(* Logix 5000 project; controller TFF vendor 1 type 14 code 107 rev 34.11; software revision 34.03; part 11 of 36 *)

        [5,29].Action := -999, [5,29].Label := -999, [5,29].Criteria1Value := -1000000.0, [5,29].Criteria2Value := -1000000.0, [5,29].ActionValue := -1000000.0, [5,30].Criteria1 := -999, [5,30].Criteria1Operator := -999, [5,30].Boolean := -999, [5,30].Criteria2 := -999, [5,30].Criteria2Operator := -999, [5,30].Action := -999, [5,30].Label := -999, [5,30].Criteria1Value := -1000000.0, [5,30].Criteria2Value := -1000000.0, [5,30].ActionValue := -1000000.0, [5,31].Criteria1 := -999, [5,31].Criteria1Operator := -999, [5,31].Boolean := -999, [5,31].Criteria2 := -999, [5,31].Criteria2Operator := -999, [5,31].Action := -999, [5,31].Label := -999, [5,31].Criteria1Value := -1000000.0, [5,31].Criteria2Value := -1000000.0, [5,31].ActionValue := -1000000.0, [5,32].Criteria1 := -999, [5,32].Criteria1Operator := -999, [5,32].Boolean := -999, [5,32].Criteria2 := -999, [5,32].Criteria2Operator := -999, [5,32].Action := -999, [5,32].Label := -999, [5,32].Criteria1Value := -1000000.0, [5,32].Criteria2Value := -1000000.0, [5,32].ActionValue := -1000000.0, [5,33].Criteria1 := -999, [5,33].Criteria1Operator := -999, [5,33].Boolean := -999, [5,33].Criteria2 := -999, [5,33].Criteria2Operator := -999, [5,33].Action := -999, [5,33].Label := -999, [5,33].Criteria1Value := -1000000.0, [5,33].Criteria2Value := -1000000.0, [5,33].ActionValue := -1000000.0, [5,34].Criteria1 := -999, [5,34].Criteria1Operator := -999, [5,34].Boolean := -999, [5,34].Criteria2 := -999, [5,34].Criteria2Operator := -999, [5,34].Action := -999, [5,34].Label := -999, [5,34].Criteria1Value := -1000000.0, [5,34].Criteria2Value := -1000000.0, [5,34].ActionValue := -1000000.0, [5,35].Criteria1 := -999, [5,35].Criteria1Operator := -999, [5,35].Boolean := -999, [5,35].Criteria2 := -999, [5,35].Criteria2Operator := -999,
        [5,35].Action := -999, [5,35].Label := -999, [5,35].Criteria1Value := -1000000.0, [5,35].Criteria2Value := -1000000.0, [5,35].ActionValue := -1000000.0, [5,36].Criteria1 := -999, [5,36].Criteria1Operator := -999, [5,36].Boolean := -999, [5,36].Criteria2 := -999, [5,36].Criteria2Operator := -999, [5,36].Action := -999, [5,36].Label := -999, [5,36].Criteria1Value := -1000000.0, [5,36].Criteria2Value := -1000000.0, [5,36].ActionValue := -1000000.0, [5,37].Criteria1 := -999, [5,37].Criteria1Operator := -999, [5,37].Boolean := -999, [5,37].Criteria2 := -999, [5,37].Criteria2Operator := -999, [5,37].Action := -999, [5,37].Label := -999, [5,37].Criteria1Value := -1000000.0, [5,37].Criteria2Value := -1000000.0, [5,37].ActionValue := -1000000.0, [5,38].Criteria1 := -999, [5,38].Criteria1Operator := -999, [5,38].Boolean := -999, [5,38].Criteria2 := -999, [5,38].Criteria2Operator := -999, [5,38].Action := -999, [5,38].Label := -999, [5,38].Criteria1Value := -1000000.0, [5,38].Criteria2Value := -1000000.0, [5,38].ActionValue := -1000000.0, [5,39].Criteria1 := -999, [5,39].Criteria1Operator := -999, [5,39].Boolean := -999, [5,39].Criteria2 := -999, [5,39].Criteria2Operator := -999, [5,39].Action := -999, [5,39].Label := -999, [5,39].Criteria1Value := -1000000.0, [5,39].Criteria2Value := -1000000.0, [5,39].ActionValue := -1000000.0, [5,40].Criteria1 := -999, [5,40].Criteria1Operator := -999, [5,40].Boolean := -999, [5,40].Criteria2 := -999, [5,40].Criteria2Operator := -999, [5,40].Action := -999, [5,40].Label := -999, [5,40].Criteria1Value := -1000000.0, [5,40].Criteria2Value := -1000000.0, [5,40].ActionValue := -1000000.0, [5,41].Criteria1 := -999, [5,41].Criteria1Operator := -999, [5,41].Boolean := -999, [5,41].Criteria2 := -999, [5,41].Criteria2Operator := -999,
        [5,41].Action := -999, [5,41].Label := -999, [5,41].Criteria1Value := -1000000.0, [5,41].Criteria2Value := -1000000.0, [5,41].ActionValue := -1000000.0, [5,42].Criteria1 := -999, [5,42].Criteria1Operator := -999, [5,42].Boolean := -999, [5,42].Criteria2 := -999, [5,42].Criteria2Operator := -999, [5,42].Action := -999, [5,42].Label := -999, [5,42].Criteria1Value := -1000000.0, [5,42].Criteria2Value := -1000000.0, [5,42].ActionValue := -1000000.0, [5,43].Criteria1 := -999, [5,43].Criteria1Operator := -999, [5,43].Boolean := -999, [5,43].Criteria2 := -999, [5,43].Criteria2Operator := -999, [5,43].Action := -999, [5,43].Label := -999, [5,43].Criteria1Value := -1000000.0, [5,43].Criteria2Value := -1000000.0, [5,43].ActionValue := -1000000.0, [5,44].Criteria1 := -999, [5,44].Criteria1Operator := -999, [5,44].Boolean := -999, [5,44].Criteria2 := -999, [5,44].Criteria2Operator := -999, [5,44].Action := -999, [5,44].Label := -999, [5,44].Criteria1Value := -1000000.0, [5,44].Criteria2Value := -1000000.0, [5,44].ActionValue := -1000000.0, [5,45].Criteria1 := -999, [5,45].Criteria1Operator := -999, [5,45].Boolean := -999, [5,45].Criteria2 := -999, [5,45].Criteria2Operator := -999, [5,45].Action := -999, [5,45].Label := -999, [5,45].Criteria1Value := -1000000.0, [5,45].Criteria2Value := -1000000.0, [5,45].ActionValue := -1000000.0, [5,46].Criteria1 := -999, [5,46].Criteria1Operator := -999, [5,46].Boolean := -999, [5,46].Criteria2 := -999, [5,46].Criteria2Operator := -999, [5,46].Action := -999, [5,46].Label := -999, [5,46].Criteria1Value := -1000000.0, [5,46].Criteria2Value := -1000000.0, [5,46].ActionValue := -1000000.0, [5,47].Criteria1 := -999, [5,47].Criteria1Operator := -999, [5,47].Boolean := -999, [5,47].Criteria2 := -999, [5,47].Criteria2Operator := -999,
        [5,47].Action := -999, [5,47].Label := -999, [5,47].Criteria1Value := -1000000.0, [5,47].Criteria2Value := -1000000.0, [5,47].ActionValue := -1000000.0, [5,48].Criteria1 := -999, [5,48].Criteria1Operator := -999, [5,48].Boolean := -999, [5,48].Criteria2 := -999, [5,48].Criteria2Operator := -999, [5,48].Action := -999, [5,48].Label := -999, [5,48].Criteria1Value := -1000000.0, [5,48].Criteria2Value := -1000000.0, [5,48].ActionValue := -1000000.0, [5,49].Criteria1 := -999, [5,49].Criteria1Operator := -999, [5,49].Boolean := -999, [5,49].Criteria2 := -999, [5,49].Criteria2Operator := -999, [5,49].Action := -999, [5,49].Label := -999, [5,49].Criteria1Value := -1000000.0, [5,49].Criteria2Value := -1000000.0, [5,49].ActionValue := -1000000.0, [5,50].Criteria1 := -999, [5,50].Criteria1Operator := -999, [5,50].Boolean := -999, [5,50].Criteria2 := -999, [5,50].Criteria2Operator := -999, [5,50].Action := -999, [5,50].Label := -999, [5,50].Criteria1Value := -1000000.0, [5,50].Criteria2Value := -1000000.0, [5,50].ActionValue := -1000000.0, [5,51].Criteria1 := -999, [5,51].Criteria1Operator := -999, [5,51].Boolean := -999, [5,51].Criteria2 := -999, [5,51].Criteria2Operator := -999, [5,51].Action := -999, [5,51].Label := -999, [5,51].Criteria1Value := -1000000.0, [5,51].Criteria2Value := -1000000.0, [5,51].ActionValue := -1000000.0, [5,52].Criteria1 := -999, [5,52].Criteria1Operator := -999, [5,52].Boolean := -999, [5,52].Criteria2 := -999, [5,52].Criteria2Operator := -999, [5,52].Action := -999, [5,52].Label := -999, [5,52].Criteria1Value := -1000000.0, [5,52].Criteria2Value := -1000000.0, [5,52].ActionValue := -1000000.0, [5,53].Criteria1 := -999, [5,53].Criteria1Operator := -999, [5,53].Boolean := -999, [5,53].Criteria2 := -999, [5,53].Criteria2Operator := -999,
        [5,53].Action := -999, [5,53].Label := -999, [5,53].Criteria1Value := -1000000.0, [5,53].Criteria2Value := -1000000.0, [5,53].ActionValue := -1000000.0, [5,54].Criteria1 := -999, [5,54].Criteria1Operator := -999, [5,54].Boolean := -999, [5,54].Criteria2 := -999, [5,54].Criteria2Operator := -999, [5,54].Action := -999, [5,54].Label := -999, [5,54].Criteria1Value := -1000000.0, [5,54].Criteria2Value := -1000000.0, [5,54].ActionValue := -1000000.0, [5,55].Criteria1 := -999, [5,55].Criteria1Operator := -999, [5,55].Boolean := -999, [5,55].Criteria2 := -999, [5,55].Criteria2Operator := -999, [5,55].Action := -999, [5,55].Label := -999, [5,55].Criteria1Value := -1000000.0, [5,55].Criteria2Value := -1000000.0, [5,55].ActionValue := -1000000.0, [5,56].Criteria1 := -999, [5,56].Criteria1Operator := -999, [5,56].Boolean := -999, [5,56].Criteria2 := -999, [5,56].Criteria2Operator := -999, [5,56].Action := -999, [5,56].Label := -999, [5,56].Criteria1Value := -1000000.0, [5,56].Criteria2Value := -1000000.0, [5,56].ActionValue := -1000000.0, [5,57].Criteria1 := -999, [5,57].Criteria1Operator := -999, [5,57].Boolean := -999, [5,57].Criteria2 := -999, [5,57].Criteria2Operator := -999, [5,57].Action := -999, [5,57].Label := -999, [5,57].Criteria1Value := -1000000.0, [5,57].Criteria2Value := -1000000.0, [5,57].ActionValue := -1000000.0, [5,58].Criteria1 := -999, [5,58].Criteria1Operator := -999, [5,58].Boolean := -999, [5,58].Criteria2 := -999, [5,58].Criteria2Operator := -999, [5,58].Action := -999, [5,58].Label := -999, [5,58].Criteria1Value := -1000000.0, [5,58].Criteria2Value := -1000000.0, [5,58].ActionValue := -1000000.0, [5,59].Criteria1 := -999, [5,59].Criteria1Operator := -999, [5,59].Boolean := -999, [5,59].Criteria2 := -999, [5,59].Criteria2Operator := -999,
        [5,59].Action := -999, [5,59].Label := -999, [5,59].Criteria1Value := -1000000.0, [5,59].Criteria2Value := -1000000.0, [5,59].ActionValue := -1000000.0, [5,60].Criteria1 := -999, [5,60].Criteria1Operator := -999, [5,60].Boolean := -999, [5,60].Criteria2 := -999, [5,60].Criteria2Operator := -999, [5,60].Action := -999, [5,60].Label := -999, [5,60].Criteria1Value := -1000000.0, [5,60].Criteria2Value := -1000000.0, [5,60].ActionValue := -1000000.0, [5,61].Criteria1 := -999, [5,61].Criteria1Operator := -999, [5,61].Boolean := -999, [5,61].Criteria2 := -999, [5,61].Criteria2Operator := -999, [5,61].Action := -999, [5,61].Label := -999, [5,61].Criteria1Value := -1000000.0, [5,61].Criteria2Value := -1000000.0, [5,61].ActionValue := -1000000.0, [5,62].Criteria1 := -999, [5,62].Criteria1Operator := -999, [5,62].Boolean := -999, [5,62].Criteria2 := -999, [5,62].Criteria2Operator := -999, [5,62].Action := -999, [5,62].Label := -999, [5,62].Criteria1Value := -1000000.0, [5,62].Criteria2Value := -1000000.0, [5,62].ActionValue := -1000000.0, [5,63].Criteria1 := -999, [5,63].Criteria1Operator := -999, [5,63].Boolean := -999, [5,63].Criteria2 := -999, [5,63].Criteria2Operator := -999, [5,63].Action := -999, [5,63].Label := -999, [5,63].Criteria1Value := -1000000.0, [5,63].Criteria2Value := -1000000.0, [5,63].ActionValue := -1000000.0, [5,64].Criteria1 := -999, [5,64].Criteria1Operator := -999, [5,64].Boolean := -999, [5,64].Criteria2 := -999, [5,64].Criteria2Operator := -999, [5,64].Action := -999, [5,64].Label := -999, [5,64].Criteria1Value := -1000000.0, [5,64].Criteria2Value := -1000000.0, [5,64].ActionValue := -1000000.0, [5,65].Criteria1 := -999, [5,65].Criteria1Operator := -999, [5,65].Boolean := -999, [5,65].Criteria2 := -999, [5,65].Criteria2Operator := -999,
        [5,65].Action := -999, [5,65].Label := -999, [5,65].Criteria1Value := -1000000.0, [5,65].Criteria2Value := -1000000.0, [5,65].ActionValue := -1000000.0, [5,66].Criteria1 := -999, [5,66].Criteria1Operator := -999, [5,66].Boolean := -999, [5,66].Criteria2 := -999, [5,66].Criteria2Operator := -999, [5,66].Action := -999, [5,66].Label := -999, [5,66].Criteria1Value := -1000000.0, [5,66].Criteria2Value := -1000000.0, [5,66].ActionValue := -1000000.0, [5,67].Criteria1 := -999, [5,67].Criteria1Operator := -999, [5,67].Boolean := -999, [5,67].Criteria2 := -999, [5,67].Criteria2Operator := -999, [5,67].Action := -999, [5,67].Label := -999, [5,67].Criteria1Value := -1000000.0, [5,67].Criteria2Value := -1000000.0, [5,67].ActionValue := -1000000.0, [5,68].Criteria1 := -999, [5,68].Criteria1Operator := -999, [5,68].Boolean := -999, [5,68].Criteria2 := -999, [5,68].Criteria2Operator := -999, [5,68].Action := -999, [5,68].Label := -999, [5,68].Criteria1Value := -1000000.0, [5,68].Criteria2Value := -1000000.0, [5,68].ActionValue := -1000000.0, [5,69].Criteria1 := -999, [5,69].Criteria1Operator := -999, [5,69].Boolean := -999, [5,69].Criteria2 := -999, [5,69].Criteria2Operator := -999, [5,69].Action := -999, [5,69].Label := -999, [5,69].Criteria1Value := -1000000.0, [5,69].Criteria2Value := -1000000.0, [5,69].ActionValue := -1000000.0, [5,70].Criteria1 := -999, [5,70].Criteria1Operator := -999, [5,70].Boolean := -999, [5,70].Criteria2 := -999, [5,70].Criteria2Operator := -999, [5,70].Action := -999, [5,70].Label := -999, [5,70].Criteria1Value := -1000000.0, [5,70].Criteria2Value := -1000000.0, [5,70].ActionValue := -1000000.0, [5,71].Criteria1 := -999, [5,71].Criteria1Operator := -999, [5,71].Boolean := -999, [5,71].Criteria2 := -999, [5,71].Criteria2Operator := -999,
        [5,71].Action := -999, [5,71].Label := -999, [5,71].Criteria1Value := -1000000.0, [5,71].Criteria2Value := -1000000.0, [5,71].ActionValue := -1000000.0, [5,72].Criteria1 := -999, [5,72].Criteria1Operator := -999, [5,72].Boolean := -999, [5,72].Criteria2 := -999, [5,72].Criteria2Operator := -999, [5,72].Action := -999, [5,72].Label := -999, [5,72].Criteria1Value := -1000000.0, [5,72].Criteria2Value := -1000000.0, [5,72].ActionValue := -1000000.0, [5,73].Criteria1 := -999, [5,73].Criteria1Operator := -999, [5,73].Boolean := -999, [5,73].Criteria2 := -999, [5,73].Criteria2Operator := -999, [5,73].Action := -999, [5,73].Label := -999, [5,73].Criteria1Value := -1000000.0, [5,73].Criteria2Value := -1000000.0, [5,73].ActionValue := -1000000.0, [5,74].Criteria1 := -999, [5,74].Criteria1Operator := -999, [5,74].Boolean := -999, [5,74].Criteria2 := -999, [5,74].Criteria2Operator := -999, [5,74].Action := -999, [5,74].Label := -999, [5,74].Criteria1Value := -1000000.0, [5,74].Criteria2Value := -1000000.0, [5,74].ActionValue := -1000000.0, [5,75].Criteria1 := -999, [5,75].Criteria1Operator := -999, [5,75].Boolean := -999, [5,75].Criteria2 := -999, [5,75].Criteria2Operator := -999, [5,75].Action := -999, [5,75].Label := -999, [5,75].Criteria1Value := -1000000.0, [5,75].Criteria2Value := -1000000.0, [5,75].ActionValue := -1000000.0, [5,76].Criteria1 := -999, [5,76].Criteria1Operator := -999, [5,76].Boolean := -999, [5,76].Criteria2 := -999, [5,76].Criteria2Operator := -999, [5,76].Action := -999, [5,76].Label := -999, [5,76].Criteria1Value := -1000000.0, [5,76].Criteria2Value := -1000000.0, [5,76].ActionValue := -1000000.0, [5,77].Criteria1 := -999, [5,77].Criteria1Operator := -999, [5,77].Boolean := -999, [5,77].Criteria2 := -999, [5,77].Criteria2Operator := -999,
        [5,77].Action := -999, [5,77].Label := -999, [5,77].Criteria1Value := -1000000.0, [5,77].Criteria2Value := -1000000.0, [5,77].ActionValue := -1000000.0, [5,78].Criteria1 := -999, [5,78].Criteria1Operator := -999, [5,78].Boolean := -999, [5,78].Criteria2 := -999, [5,78].Criteria2Operator := -999, [5,78].Action := -999, [5,78].Label := -999, [5,78].Criteria1Value := -1000000.0, [5,78].Criteria2Value := -1000000.0, [5,78].ActionValue := -1000000.0, [5,79].Criteria1 := -999, [5,79].Criteria1Operator := -999, [5,79].Boolean := -999, [5,79].Criteria2 := -999, [5,79].Criteria2Operator := -999, [5,79].Action := -999, [5,79].Label := -999, [5,79].Criteria1Value := -1000000.0, [5,79].Criteria2Value := -1000000.0, [5,79].ActionValue := -1000000.0, [5,80].Criteria1 := -999, [5,80].Criteria1Operator := -999, [5,80].Boolean := -999, [5,80].Criteria2 := -999, [5,80].Criteria2Operator := -999, [5,80].Action := -999, [5,80].Label := -999, [5,80].Criteria1Value := -1000000.0, [5,80].Criteria2Value := -1000000.0, [5,80].ActionValue := -1000000.0, [5,81].Criteria1 := -999, [5,81].Criteria1Operator := -999, [5,81].Boolean := -999, [5,81].Criteria2 := -999, [5,81].Criteria2Operator := -999, [5,81].Action := -999, [5,81].Label := -999, [5,81].Criteria1Value := -1000000.0, [5,81].Criteria2Value := -1000000.0, [5,81].ActionValue := -1000000.0, [5,82].Criteria1 := -999, [5,82].Criteria1Operator := -999, [5,82].Boolean := -999, [5,82].Criteria2 := -999, [5,82].Criteria2Operator := -999, [5,82].Action := -999, [5,82].Label := -999, [5,82].Criteria1Value := -1000000.0, [5,82].Criteria2Value := -1000000.0, [5,82].ActionValue := -1000000.0, [5,83].Criteria1 := -999, [5,83].Criteria1Operator := -999, [5,83].Boolean := -999, [5,83].Criteria2 := -999, [5,83].Criteria2Operator := -999,
        [5,83].Action := -999, [5,83].Label := -999, [5,83].Criteria1Value := -1000000.0, [5,83].Criteria2Value := -1000000.0, [5,83].ActionValue := -1000000.0, [5,84].Criteria1 := -999, [5,84].Criteria1Operator := -999, [5,84].Boolean := -999, [5,84].Criteria2 := -999, [5,84].Criteria2Operator := -999, [5,84].Action := -999, [5,84].Label := -999, [5,84].Criteria1Value := -1000000.0, [5,84].Criteria2Value := -1000000.0, [5,84].ActionValue := -1000000.0, [5,85].Criteria1 := -999, [5,85].Criteria1Operator := -999, [5,85].Boolean := -999, [5,85].Criteria2 := -999, [5,85].Criteria2Operator := -999, [5,85].Action := -999, [5,85].Label := -999, [5,85].Criteria1Value := -1000000.0, [5,85].Criteria2Value := -1000000.0, [5,85].ActionValue := -1000000.0, [5,86].Criteria1 := -999, [5,86].Criteria1Operator := -999, [5,86].Boolean := -999, [5,86].Criteria2 := -999, [5,86].Criteria2Operator := -999, [5,86].Action := -999, [5,86].Label := -999, [5,86].Criteria1Value := -1000000.0, [5,86].Criteria2Value := -1000000.0, [5,86].ActionValue := -1000000.0, [5,87].Criteria1 := -999, [5,87].Criteria1Operator := -999, [5,87].Boolean := -999, [5,87].Criteria2 := -999, [5,87].Criteria2Operator := -999, [5,87].Action := -999, [5,87].Label := -999, [5,87].Criteria1Value := -1000000.0, [5,87].Criteria2Value := -1000000.0, [5,87].ActionValue := -1000000.0, [5,88].Criteria1 := -999, [5,88].Criteria1Operator := -999, [5,88].Boolean := -999, [5,88].Criteria2 := -999, [5,88].Criteria2Operator := -999, [5,88].Action := -999, [5,88].Label := -999, [5,88].Criteria1Value := -1000000.0, [5,88].Criteria2Value := -1000000.0, [5,88].ActionValue := -1000000.0, [5,89].Criteria1 := -999, [5,89].Criteria1Operator := -999, [5,89].Boolean := -999, [5,89].Criteria2 := -999, [5,89].Criteria2Operator := -999,
        [5,89].Action := -999, [5,89].Label := -999, [5,89].Criteria1Value := -1000000.0, [5,89].Criteria2Value := -1000000.0, [5,89].ActionValue := -1000000.0, [5,90].Criteria1 := -999, [5,90].Criteria1Operator := -999, [5,90].Boolean := -999, [5,90].Criteria2 := -999, [5,90].Criteria2Operator := -999, [5,90].Action := -999, [5,90].Label := -999, [5,90].Criteria1Value := -1000000.0, [5,90].Criteria2Value := -1000000.0, [5,90].ActionValue := -1000000.0, [5,91].Criteria1 := -999, [5,91].Criteria1Operator := -999, [5,91].Boolean := -999, [5,91].Criteria2 := -999, [5,91].Criteria2Operator := -999, [5,91].Action := -999, [5,91].Label := -999, [5,91].Criteria1Value := -1000000.0, [5,91].Criteria2Value := -1000000.0, [5,91].ActionValue := -1000000.0, [5,92].Criteria1 := -999, [5,92].Criteria1Operator := -999, [5,92].Boolean := -999, [5,92].Criteria2 := -999, [5,92].Criteria2Operator := -999, [5,92].Action := -999, [5,92].Label := -999, [5,92].Criteria1Value := -1000000.0, [5,92].Criteria2Value := -1000000.0, [5,92].ActionValue := -1000000.0, [5,93].Criteria1 := -999, [5,93].Criteria1Operator := -999, [5,93].Boolean := -999, [5,93].Criteria2 := -999, [5,93].Criteria2Operator := -999, [5,93].Action := -999, [5,93].Label := -999, [5,93].Criteria1Value := -1000000.0, [5,93].Criteria2Value := -1000000.0, [5,93].ActionValue := -1000000.0, [5,94].Criteria1 := -999, [5,94].Criteria1Operator := -999, [5,94].Boolean := -999, [5,94].Criteria2 := -999, [5,94].Criteria2Operator := -999, [5,94].Action := -999, [5,94].Label := -999, [5,94].Criteria1Value := -1000000.0, [5,94].Criteria2Value := -1000000.0, [5,94].ActionValue := -1000000.0, [5,95].Criteria1 := -999, [5,95].Criteria1Operator := -999, [5,95].Boolean := -999, [5,95].Criteria2 := -999, [5,95].Criteria2Operator := -999,
        [5,95].Action := -999, [5,95].Label := -999, [5,95].Criteria1Value := -1000000.0, [5,95].Criteria2Value := -1000000.0, [5,95].ActionValue := -1000000.0, [5,96].Criteria1 := -999, [5,96].Criteria1Operator := -999, [5,96].Boolean := -999, [5,96].Criteria2 := -999, [5,96].Criteria2Operator := -999, [5,96].Action := -999, [5,96].Label := -999, [5,96].Criteria1Value := -1000000.0, [5,96].Criteria2Value := -1000000.0, [5,96].ActionValue := -1000000.0, [5,97].Criteria1 := -999, [5,97].Criteria1Operator := -999, [5,97].Boolean := -999, [5,97].Criteria2 := -999, [5,97].Criteria2Operator := -999, [5,97].Action := -999, [5,97].Label := -999, [5,97].Criteria1Value := -1000000.0, [5,97].Criteria2Value := -1000000.0, [5,97].ActionValue := -1000000.0, [5,98].Criteria1 := -999, [5,98].Criteria1Operator := -999, [5,98].Boolean := -999, [5,98].Criteria2 := -999, [5,98].Criteria2Operator := -999, [5,98].Action := -999, [5,98].Label := -999, [5,98].Criteria1Value := -1000000.0, [5,98].Criteria2Value := -1000000.0, [5,98].ActionValue := -1000000.0, [5,99].Criteria1 := -999, [5,99].Criteria1Operator := -999, [5,99].Boolean := -999, [5,99].Criteria2 := -999, [5,99].Criteria2Operator := -999, [5,99].Action := -999, [5,99].Label := -999, [5,99].Criteria1Value := -1000000.0, [5,99].Criteria2Value := -1000000.0, [5,99].ActionValue := -1000000.0, [5,100].Criteria1 := -999, [5,100].Criteria1Operator := -999, [5,100].Boolean := -999, [5,100].Criteria2 := -999, [5,100].Criteria2Operator := -999, [5,100].Action := -999, [5,100].Label := -999, [5,100].Criteria1Value := -1000000.0, [5,100].Criteria2Value := -1000000.0, [5,100].ActionValue := -1000000.0, [5,101].Criteria1 := -999, [5,101].Criteria1Operator := -999, [5,101].Boolean := -999, [5,101].Criteria2 := -999, [5,101].Criteria2Operator := -999,
        [5,101].Action := -999, [5,101].Label := -999, [5,101].Criteria1Value := -1000000.0, [5,101].Criteria2Value := -1000000.0, [5,101].ActionValue := -1000000.0, [5,102].Criteria1 := -999, [5,102].Criteria1Operator := -999, [5,102].Boolean := -999, [5,102].Criteria2 := -999, [5,102].Criteria2Operator := -999, [5,102].Action := -999, [5,102].Label := -999, [5,102].Criteria1Value := -1000000.0, [5,102].Criteria2Value := -1000000.0, [5,102].ActionValue := -1000000.0, [5,103].Criteria1 := -999, [5,103].Criteria1Operator := -999, [5,103].Boolean := -999, [5,103].Criteria2 := -999, [5,103].Criteria2Operator := -999, [5,103].Action := -999, [5,103].Label := -999, [5,103].Criteria1Value := -1000000.0, [5,103].Criteria2Value := -1000000.0, [5,103].ActionValue := -1000000.0, [5,104].Criteria1 := -999, [5,104].Criteria1Operator := -999, [5,104].Boolean := -999, [5,104].Criteria2 := -999, [5,104].Criteria2Operator := -999, [5,104].Action := -999, [5,104].Label := -999, [5,104].Criteria1Value := -1000000.0, [5,104].Criteria2Value := -1000000.0, [5,104].ActionValue := -1000000.0, [5,105].Criteria1 := -999, [5,105].Criteria1Operator := -999, [5,105].Boolean := -999, [5,105].Criteria2 := -999, [5,105].Criteria2Operator := -999, [5,105].Action := -999, [5,105].Label := -999, [5,105].Criteria1Value := -1000000.0, [5,105].Criteria2Value := -1000000.0, [5,105].ActionValue := -1000000.0, [5,106].Criteria1 := -999, [5,106].Criteria1Operator := -999, [5,106].Boolean := -999, [5,106].Criteria2 := -999, [5,106].Criteria2Operator := -999, [5,106].Action := -999, [5,106].Label := -999, [5,106].Criteria1Value := -1000000.0, [5,106].Criteria2Value := -1000000.0, [5,106].ActionValue := -1000000.0, [5,107].Criteria1 := -999, [5,107].Criteria1Operator := -999, [5,107].Boolean := -999, [5,107].Criteria2 := -999, [5,107].Criteria2Operator := -999,
        [5,107].Action := -999, [5,107].Label := -999, [5,107].Criteria1Value := -1000000.0, [5,107].Criteria2Value := -1000000.0, [5,107].ActionValue := -1000000.0, [5,108].Criteria1 := -999, [5,108].Criteria1Operator := -999, [5,108].Boolean := -999, [5,108].Criteria2 := -999, [5,108].Criteria2Operator := -999, [5,108].Action := -999, [5,108].Label := -999, [5,108].Criteria1Value := -1000000.0, [5,108].Criteria2Value := -1000000.0, [5,108].ActionValue := -1000000.0, [5,109].Criteria1 := -999, [5,109].Criteria1Operator := -999, [5,109].Boolean := -999, [5,109].Criteria2 := -999, [5,109].Criteria2Operator := -999, [5,109].Action := -999, [5,109].Label := -999, [5,109].Criteria1Value := -1000000.0, [5,109].Criteria2Value := -1000000.0, [5,109].ActionValue := -1000000.0, [5,110].Criteria1 := -999, [5,110].Criteria1Operator := -999, [5,110].Boolean := -999, [5,110].Criteria2 := -999, [5,110].Criteria2Operator := -999, [5,110].Action := -999, [5,110].Label := -999, [5,110].Criteria1Value := -1000000.0, [5,110].Criteria2Value := -1000000.0, [5,110].ActionValue := -1000000.0, [5,111].Criteria1 := -999, [5,111].Criteria1Operator := -999, [5,111].Boolean := -999, [5,111].Criteria2 := -999, [5,111].Criteria2Operator := -999, [5,111].Action := -999, [5,111].Label := -999, [5,111].Criteria1Value := -1000000.0, [5,111].Criteria2Value := -1000000.0, [5,111].ActionValue := -1000000.0, [5,112].Criteria1 := -999, [5,112].Criteria1Operator := -999, [5,112].Boolean := -999, [5,112].Criteria2 := -999, [5,112].Criteria2Operator := -999, [5,112].Action := -999, [5,112].Label := -999, [5,112].Criteria1Value := -1000000.0, [5,112].Criteria2Value := -1000000.0, [5,112].ActionValue := -1000000.0, [5,113].Criteria1 := -999, [5,113].Criteria1Operator := -999, [5,113].Boolean := -999, [5,113].Criteria2 := -999, [5,113].Criteria2Operator := -999,
        [5,113].Action := -999, [5,113].Label := -999, [5,113].Criteria1Value := -1000000.0, [5,113].Criteria2Value := -1000000.0, [5,113].ActionValue := -1000000.0, [5,114].Criteria1 := -999, [5,114].Criteria1Operator := -999, [5,114].Boolean := -999, [5,114].Criteria2 := -999, [5,114].Criteria2Operator := -999, [5,114].Action := -999, [5,114].Label := -999, [5,114].Criteria1Value := -1000000.0, [5,114].Criteria2Value := -1000000.0, [5,114].ActionValue := -1000000.0, [5,115].Criteria1 := -999, [5,115].Criteria1Operator := -999, [5,115].Boolean := -999, [5,115].Criteria2 := -999, [5,115].Criteria2Operator := -999, [5,115].Action := -999, [5,115].Label := -999, [5,115].Criteria1Value := -1000000.0, [5,115].Criteria2Value := -1000000.0, [5,115].ActionValue := -1000000.0, [5,116].Criteria1 := -999, [5,116].Criteria1Operator := -999, [5,116].Boolean := -999, [5,116].Criteria2 := -999, [5,116].Criteria2Operator := -999, [5,116].Action := -999, [5,116].Label := -999, [5,116].Criteria1Value := -1000000.0, [5,116].Criteria2Value := -1000000.0, [5,116].ActionValue := -1000000.0, [5,117].Criteria1 := -999, [5,117].Criteria1Operator := -999, [5,117].Boolean := -999, [5,117].Criteria2 := -999, [5,117].Criteria2Operator := -999, [5,117].Action := -999, [5,117].Label := -999, [5,117].Criteria1Value := -1000000.0, [5,117].Criteria2Value := -1000000.0, [5,117].ActionValue := -1000000.0, [5,118].Criteria1 := -999, [5,118].Criteria1Operator := -999, [5,118].Boolean := -999, [5,118].Criteria2 := -999, [5,118].Criteria2Operator := -999, [5,118].Action := -999, [5,118].Label := -999, [5,118].Criteria1Value := -1000000.0, [5,118].Criteria2Value := -1000000.0, [5,118].ActionValue := -1000000.0, [5,119].Criteria1 := -999, [5,119].Criteria1Operator := -999, [5,119].Boolean := -999, [5,119].Criteria2 := -999, [5,119].Criteria2Operator := -999,
        [5,119].Action := -999, [5,119].Label := -999, [5,119].Criteria1Value := -1000000.0, [5,119].Criteria2Value := -1000000.0, [5,119].ActionValue := -1000000.0, [5,120].Criteria1 := -999, [5,120].Criteria1Operator := -999, [5,120].Boolean := -999, [5,120].Criteria2 := -999, [5,120].Criteria2Operator := -999, [5,120].Action := -999, [5,120].Label := -999, [5,120].Criteria1Value := -1000000.0, [5,120].Criteria2Value := -1000000.0, [5,120].ActionValue := -1000000.0, [5,121].Criteria1 := -999, [5,121].Criteria1Operator := -999, [5,121].Boolean := -999, [5,121].Criteria2 := -999, [5,121].Criteria2Operator := -999, [5,121].Action := -999, [5,121].Label := -999, [5,121].Criteria1Value := -1000000.0, [5,121].Criteria2Value := -1000000.0, [5,121].ActionValue := -1000000.0, [5,122].Criteria1 := -999, [5,122].Criteria1Operator := -999, [5,122].Boolean := -999, [5,122].Criteria2 := -999, [5,122].Criteria2Operator := -999, [5,122].Action := -999, [5,122].Label := -999, [5,122].Criteria1Value := -1000000.0, [5,122].Criteria2Value := -1000000.0, [5,122].ActionValue := -1000000.0, [5,123].Criteria1 := -999, [5,123].Criteria1Operator := -999, [5,123].Boolean := -999, [5,123].Criteria2 := -999, [5,123].Criteria2Operator := -999, [5,123].Action := -999, [5,123].Label := -999, [5,123].Criteria1Value := -1000000.0, [5,123].Criteria2Value := -1000000.0, [5,123].ActionValue := -1000000.0, [5,124].Criteria1 := -999, [5,124].Criteria1Operator := -999, [5,124].Boolean := -999, [5,124].Criteria2 := -999, [5,124].Criteria2Operator := -999, [5,124].Action := -999, [5,124].Label := -999, [5,124].Criteria1Value := -1000000.0, [5,124].Criteria2Value := -1000000.0, [5,124].ActionValue := -1000000.0, [5,125].Criteria1 := -999, [5,125].Criteria1Operator := -999, [5,125].Boolean := -999, [5,125].Criteria2 := -999, [5,125].Criteria2Operator := -999,
        [5,125].Action := -999, [5,125].Label := -999, [5,125].Criteria1Value := -1000000.0, [5,125].Criteria2Value := -1000000.0, [5,125].ActionValue := -1000000.0, [5,126].Criteria1 := -999, [5,126].Criteria1Operator := -999, [5,126].Boolean := -999, [5,126].Criteria2 := -999, [5,126].Criteria2Operator := -999, [5,126].Action := -999, [5,126].Label := -999, [5,126].Criteria1Value := -1000000.0, [5,126].Criteria2Value := -1000000.0, [5,126].ActionValue := -1000000.0, [5,127].Criteria1 := -999, [5,127].Criteria1Operator := -999, [5,127].Boolean := -999, [5,127].Criteria2 := -999, [5,127].Criteria2Operator := -999, [5,127].Action := -999, [5,127].Label := -999, [5,127].Criteria1Value := -1000000.0, [5,127].Criteria2Value := -1000000.0, [5,127].ActionValue := -1000000.0, [5,128].Criteria1 := -999, [5,128].Criteria1Operator := -999, [5,128].Boolean := -999, [5,128].Criteria2 := -999, [5,128].Criteria2Operator := -999, [5,128].Action := -999, [5,128].Label := -999, [5,128].Criteria1Value := -1000000.0, [5,128].Criteria2Value := -1000000.0, [5,128].ActionValue := -1000000.0, [5,129].Criteria1 := -999, [5,129].Criteria1Operator := -999, [5,129].Boolean := -999, [5,129].Criteria2 := -999, [5,129].Criteria2Operator := -999, [5,129].Action := -999, [5,129].Label := -999, [5,129].Criteria1Value := -1000000.0, [5,129].Criteria2Value := -1000000.0, [5,129].ActionValue := -1000000.0, [5,130].Criteria1 := -999, [5,130].Criteria1Operator := -999, [5,130].Boolean := -999, [5,130].Criteria2 := -999, [5,130].Criteria2Operator := -999, [5,130].Action := -999, [5,130].Label := -999, [5,130].Criteria1Value := -1000000.0, [5,130].Criteria2Value := -1000000.0, [5,130].ActionValue := -1000000.0, [5,131].Criteria1 := -999, [5,131].Criteria1Operator := -999, [5,131].Boolean := -999, [5,131].Criteria2 := -999, [5,131].Criteria2Operator := -999,
        [5,131].Action := -999, [5,131].Label := -999, [5,131].Criteria1Value := -1000000.0, [5,131].Criteria2Value := -1000000.0, [5,131].ActionValue := -1000000.0, [5,132].Criteria1 := -999, [5,132].Criteria1Operator := -999, [5,132].Boolean := -999, [5,132].Criteria2 := -999, [5,132].Criteria2Operator := -999, [5,132].Action := -999, [5,132].Label := -999, [5,132].Criteria1Value := -1000000.0, [5,132].Criteria2Value := -1000000.0, [5,132].ActionValue := -1000000.0, [5,133].Criteria1 := -999, [5,133].Criteria1Operator := -999, [5,133].Boolean := -999, [5,133].Criteria2 := -999, [5,133].Criteria2Operator := -999, [5,133].Action := -999, [5,133].Label := -999, [5,133].Criteria1Value := -1000000.0, [5,133].Criteria2Value := -1000000.0, [5,133].ActionValue := -1000000.0, [5,134].Criteria1 := -999, [5,134].Criteria1Operator := -999, [5,134].Boolean := -999, [5,134].Criteria2 := -999, [5,134].Criteria2Operator := -999, [5,134].Action := -999, [5,134].Label := -999, [5,134].Criteria1Value := -1000000.0, [5,134].Criteria2Value := -1000000.0, [5,134].ActionValue := -1000000.0, [5,135].Criteria1 := -999, [5,135].Criteria1Operator := -999, [5,135].Boolean := -999, [5,135].Criteria2 := -999, [5,135].Criteria2Operator := -999, [5,135].Action := -999, [5,135].Label := -999, [5,135].Criteria1Value := -1000000.0, [5,135].Criteria2Value := -1000000.0, [5,135].ActionValue := -1000000.0, [5,136].Criteria1 := -999, [5,136].Criteria1Operator := -999, [5,136].Boolean := -999, [5,136].Criteria2 := -999, [5,136].Criteria2Operator := -999, [5,136].Action := -999, [5,136].Label := -999, [5,136].Criteria1Value := -1000000.0, [5,136].Criteria2Value := -1000000.0, [5,136].ActionValue := -1000000.0, [5,137].Criteria1 := -999, [5,137].Criteria1Operator := -999, [5,137].Boolean := -999, [5,137].Criteria2 := -999, [5,137].Criteria2Operator := -999,
        [5,137].Action := -999, [5,137].Label := -999, [5,137].Criteria1Value := -1000000.0, [5,137].Criteria2Value := -1000000.0, [5,137].ActionValue := -1000000.0, [5,138].Criteria1 := -999, [5,138].Criteria1Operator := -999, [5,138].Boolean := -999, [5,138].Criteria2 := -999, [5,138].Criteria2Operator := -999, [5,138].Action := -999, [5,138].Label := -999, [5,138].Criteria1Value := -1000000.0, [5,138].Criteria2Value := -1000000.0, [5,138].ActionValue := -1000000.0, [5,139].Criteria1 := -999, [5,139].Criteria1Operator := -999, [5,139].Boolean := -999, [5,139].Criteria2 := -999, [5,139].Criteria2Operator := -999, [5,139].Action := -999, [5,139].Label := -999, [5,139].Criteria1Value := -1000000.0, [5,139].Criteria2Value := -1000000.0, [5,139].ActionValue := -1000000.0, [5,140].Criteria1 := -999, [5,140].Criteria1Operator := -999, [5,140].Boolean := -999, [5,140].Criteria2 := -999, [5,140].Criteria2Operator := -999, [5,140].Action := -999, [5,140].Label := -999, [5,140].Criteria1Value := -1000000.0, [5,140].Criteria2Value := -1000000.0, [5,140].ActionValue := -1000000.0, [5,141].Criteria1 := -999, [5,141].Criteria1Operator := -999, [5,141].Boolean := -999, [5,141].Criteria2 := -999, [5,141].Criteria2Operator := -999, [5,141].Action := -999, [5,141].Label := -999, [5,141].Criteria1Value := -1000000.0, [5,141].Criteria2Value := -1000000.0, [5,141].ActionValue := -1000000.0, [5,142].Criteria1 := -999, [5,142].Criteria1Operator := -999, [5,142].Boolean := -999, [5,142].Criteria2 := -999, [5,142].Criteria2Operator := -999, [5,142].Action := -999, [5,142].Label := -999, [5,142].Criteria1Value := -1000000.0, [5,142].Criteria2Value := -1000000.0, [5,142].ActionValue := -1000000.0, [5,143].Criteria1 := -999, [5,143].Criteria1Operator := -999, [5,143].Boolean := -999, [5,143].Criteria2 := -999, [5,143].Criteria2Operator := -999,
        [5,143].Action := -999, [5,143].Label := -999, [5,143].Criteria1Value := -1000000.0, [5,143].Criteria2Value := -1000000.0, [5,143].ActionValue := -1000000.0, [5,144].Criteria1 := -999, [5,144].Criteria1Operator := -999, [5,144].Boolean := -999, [5,144].Criteria2 := -999, [5,144].Criteria2Operator := -999, [5,144].Action := -999, [5,144].Label := -999, [5,144].Criteria1Value := -1000000.0, [5,144].Criteria2Value := -1000000.0, [5,144].ActionValue := -1000000.0, [5,145].Criteria1 := -999, [5,145].Criteria1Operator := -999, [5,145].Boolean := -999, [5,145].Criteria2 := -999, [5,145].Criteria2Operator := -999, [5,145].Action := -999, [5,145].Label := -999, [5,145].Criteria1Value := -1000000.0, [5,145].Criteria2Value := -1000000.0, [5,145].ActionValue := -1000000.0, [5,146].Criteria1 := -999, [5,146].Criteria1Operator := -999, [5,146].Boolean := -999, [5,146].Criteria2 := -999, [5,146].Criteria2Operator := -999, [5,146].Action := -999, [5,146].Label := -999, [5,146].Criteria1Value := -1000000.0, [5,146].Criteria2Value := -1000000.0, [5,146].ActionValue := -1000000.0, [5,147].Criteria1 := -999, [5,147].Criteria1Operator := -999, [5,147].Boolean := -999, [5,147].Criteria2 := -999, [5,147].Criteria2Operator := -999, [5,147].Action := -999, [5,147].Label := -999, [5,147].Criteria1Value := -1000000.0, [5,147].Criteria2Value := -1000000.0, [5,147].ActionValue := -1000000.0, [5,148].Criteria1 := -999, [5,148].Criteria1Operator := -999, [5,148].Boolean := -999, [5,148].Criteria2 := -999, [5,148].Criteria2Operator := -999, [5,148].Action := -999, [5,148].Label := -999, [5,148].Criteria1Value := -1000000.0, [5,148].Criteria2Value := -1000000.0, [5,148].ActionValue := -1000000.0, [5,149].Criteria1 := -999, [5,149].Criteria1Operator := -999, [5,149].Boolean := -999, [5,149].Criteria2 := -999, [5,149].Criteria2Operator := -999,
        [5,149].Action := -999, [5,149].Label := -999, [5,149].Criteria1Value := -1000000.0, [5,149].Criteria2Value := -1000000.0, [5,149].ActionValue := -1000000.0, [5,150].Criteria1 := -999, [5,150].Criteria1Operator := -999, [5,150].Boolean := -999, [5,150].Criteria2 := -999, [5,150].Criteria2Operator := -999, [5,150].Action := -999, [5,150].Label := -999, [5,150].Criteria1Value := -1000000.0, [5,150].Criteria2Value := -1000000.0, [5,150].ActionValue := -1000000.0, [5,151].Criteria1 := -999, [5,151].Criteria1Operator := -999, [5,151].Boolean := -999, [5,151].Criteria2 := -999, [5,151].Criteria2Operator := -999, [5,151].Action := -999, [5,151].Label := -999, [5,151].Criteria1Value := -1000000.0, [5,151].Criteria2Value := -1000000.0, [5,151].ActionValue := -1000000.0, [5,152].Criteria1 := -999, [5,152].Criteria1Operator := -999, [5,152].Boolean := -999, [5,152].Criteria2 := -999, [5,152].Criteria2Operator := -999, [5,152].Action := -999, [5,152].Label := -999, [5,152].Criteria1Value := -1000000.0, [5,152].Criteria2Value := -1000000.0, [5,152].ActionValue := -1000000.0, [5,153].Criteria1 := -999, [5,153].Criteria1Operator := -999, [5,153].Boolean := -999, [5,153].Criteria2 := -999, [5,153].Criteria2Operator := -999, [5,153].Action := -999, [5,153].Label := -999, [5,153].Criteria1Value := -1000000.0, [5,153].Criteria2Value := -1000000.0, [5,153].ActionValue := -1000000.0, [5,154].Criteria1 := -999, [5,154].Criteria1Operator := -999, [5,154].Boolean := -999, [5,154].Criteria2 := -999, [5,154].Criteria2Operator := -999, [5,154].Action := -999, [5,154].Label := -999, [5,154].Criteria1Value := -1000000.0, [5,154].Criteria2Value := -1000000.0, [5,154].ActionValue := -1000000.0, [5,155].Criteria1 := -999, [5,155].Criteria1Operator := -999, [5,155].Boolean := -999, [5,155].Criteria2 := -999, [5,155].Criteria2Operator := -999,
        [5,155].Action := -999, [5,155].Label := -999, [5,155].Criteria1Value := -1000000.0, [5,155].Criteria2Value := -1000000.0, [5,155].ActionValue := -1000000.0, [5,156].Criteria1 := -999, [5,156].Criteria1Operator := -999, [5,156].Boolean := -999, [5,156].Criteria2 := -999, [5,156].Criteria2Operator := -999, [5,156].Action := -999, [5,156].Label := -999, [5,156].Criteria1Value := -1000000.0, [5,156].Criteria2Value := -1000000.0, [5,156].ActionValue := -1000000.0, [5,157].Criteria1 := -999, [5,157].Criteria1Operator := -999, [5,157].Boolean := -999, [5,157].Criteria2 := -999, [5,157].Criteria2Operator := -999, [5,157].Action := -999, [5,157].Label := -999, [5,157].Criteria1Value := -1000000.0, [5,157].Criteria2Value := -1000000.0, [5,157].ActionValue := -1000000.0, [5,158].Criteria1 := -999, [5,158].Criteria1Operator := -999, [5,158].Boolean := -999, [5,158].Criteria2 := -999, [5,158].Criteria2Operator := -999, [5,158].Action := -999, [5,158].Label := -999, [5,158].Criteria1Value := -1000000.0, [5,158].Criteria2Value := -1000000.0, [5,158].ActionValue := -1000000.0, [5,159].Criteria1 := -999, [5,159].Criteria1Operator := -999, [5,159].Boolean := -999, [5,159].Criteria2 := -999, [5,159].Criteria2Operator := -999, [5,159].Action := -999, [5,159].Label := -999, [5,159].Criteria1Value := -1000000.0, [5,159].Criteria2Value := -1000000.0, [5,159].ActionValue := -1000000.0, [5,160].Criteria1 := -999, [5,160].Criteria1Operator := -999, [5,160].Boolean := -999, [5,160].Criteria2 := -999, [5,160].Criteria2Operator := -999, [5,160].Action := -999, [5,160].Label := -999, [5,160].Criteria1Value := -1000000.0, [5,160].Criteria2Value := -1000000.0, [5,160].ActionValue := -1000000.0, [5,161].Criteria1 := -999, [5,161].Criteria1Operator := -999, [5,161].Boolean := -999, [5,161].Criteria2 := -999, [5,161].Criteria2Operator := -999,
        [5,161].Action := -999, [5,161].Label := -999, [5,161].Criteria1Value := -1000000.0, [5,161].Criteria2Value := -1000000.0, [5,161].ActionValue := -1000000.0, [5,162].Criteria1 := -999, [5,162].Criteria1Operator := -999, [5,162].Boolean := -999, [5,162].Criteria2 := -999, [5,162].Criteria2Operator := -999, [5,162].Action := -999, [5,162].Label := -999, [5,162].Criteria1Value := -1000000.0, [5,162].Criteria2Value := -1000000.0, [5,162].ActionValue := -1000000.0, [5,163].Criteria1 := -999, [5,163].Criteria1Operator := -999, [5,163].Boolean := -999, [5,163].Criteria2 := -999, [5,163].Criteria2Operator := -999, [5,163].Action := -999, [5,163].Label := -999, [5,163].Criteria1Value := -1000000.0, [5,163].Criteria2Value := -1000000.0, [5,163].ActionValue := -1000000.0, [5,164].Criteria1 := -999, [5,164].Criteria1Operator := -999, [5,164].Boolean := -999, [5,164].Criteria2 := -999, [5,164].Criteria2Operator := -999, [5,164].Action := -999, [5,164].Label := -999, [5,164].Criteria1Value := -1000000.0, [5,164].Criteria2Value := -1000000.0, [5,164].ActionValue := -1000000.0, [5,165].Criteria1 := -999, [5,165].Criteria1Operator := -999, [5,165].Boolean := -999, [5,165].Criteria2 := -999, [5,165].Criteria2Operator := -999, [5,165].Action := -999, [5,165].Label := -999, [5,165].Criteria1Value := -1000000.0, [5,165].Criteria2Value := -1000000.0, [5,165].ActionValue := -1000000.0, [5,166].Criteria1 := -999, [5,166].Criteria1Operator := -999, [5,166].Boolean := -999, [5,166].Criteria2 := -999, [5,166].Criteria2Operator := -999, [5,166].Action := -999, [5,166].Label := -999, [5,166].Criteria1Value := -1000000.0, [5,166].Criteria2Value := -1000000.0, [5,166].ActionValue := -1000000.0, [5,167].Criteria1 := -999, [5,167].Criteria1Operator := -999, [5,167].Boolean := -999, [5,167].Criteria2 := -999, [5,167].Criteria2Operator := -999,
        [5,167].Action := -999, [5,167].Label := -999, [5,167].Criteria1Value := -1000000.0, [5,167].Criteria2Value := -1000000.0, [5,167].ActionValue := -1000000.0, [5,168].Criteria1 := -999, [5,168].Criteria1Operator := -999, [5,168].Boolean := -999, [5,168].Criteria2 := -999, [5,168].Criteria2Operator := -999, [5,168].Action := -999, [5,168].Label := -999, [5,168].Criteria1Value := -1000000.0, [5,168].Criteria2Value := -1000000.0, [5,168].ActionValue := -1000000.0, [5,169].Criteria1 := -999, [5,169].Criteria1Operator := -999, [5,169].Boolean := -999, [5,169].Criteria2 := -999, [5,169].Criteria2Operator := -999, [5,169].Action := -999, [5,169].Label := -999, [5,169].Criteria1Value := -1000000.0, [5,169].Criteria2Value := -1000000.0, [5,169].ActionValue := -1000000.0, [5,170].Criteria1 := -999, [5,170].Criteria1Operator := -999, [5,170].Boolean := -999, [5,170].Criteria2 := -999, [5,170].Criteria2Operator := -999, [5,170].Action := -999, [5,170].Label := -999, [5,170].Criteria1Value := -1000000.0, [5,170].Criteria2Value := -1000000.0, [5,170].ActionValue := -1000000.0, [5,171].Criteria1 := -999, [5,171].Criteria1Operator := -999, [5,171].Boolean := -999, [5,171].Criteria2 := -999, [5,171].Criteria2Operator := -999, [5,171].Action := -999, [5,171].Label := -999, [5,171].Criteria1Value := -1000000.0, [5,171].Criteria2Value := -1000000.0, [5,171].ActionValue := -1000000.0, [5,172].Criteria1 := -999, [5,172].Criteria1Operator := -999, [5,172].Boolean := -999, [5,172].Criteria2 := -999, [5,172].Criteria2Operator := -999, [5,172].Action := -999, [5,172].Label := -999, [5,172].Criteria1Value := -1000000.0, [5,172].Criteria2Value := -1000000.0, [5,172].ActionValue := -1000000.0, [5,173].Criteria1 := -999, [5,173].Criteria1Operator := -999, [5,173].Boolean := -999, [5,173].Criteria2 := -999, [5,173].Criteria2Operator := -999,
        [5,173].Action := -999, [5,173].Label := -999, [5,173].Criteria1Value := -1000000.0, [5,173].Criteria2Value := -1000000.0, [5,173].ActionValue := -1000000.0, [5,174].Criteria1 := -999, [5,174].Criteria1Operator := -999, [5,174].Boolean := -999, [5,174].Criteria2 := -999, [5,174].Criteria2Operator := -999, [5,174].Action := -999, [5,174].Label := -999, [5,174].Criteria1Value := -1000000.0, [5,174].Criteria2Value := -1000000.0, [5,174].ActionValue := -1000000.0, [5,175].Criteria1 := -999, [5,175].Criteria1Operator := -999, [5,175].Boolean := -999, [5,175].Criteria2 := -999, [5,175].Criteria2Operator := -999, [5,175].Action := -999, [5,175].Label := -999, [5,175].Criteria1Value := -1000000.0, [5,175].Criteria2Value := -1000000.0, [5,175].ActionValue := -1000000.0, [5,176].Criteria1 := -999, [5,176].Criteria1Operator := -999, [5,176].Boolean := -999, [5,176].Criteria2 := -999, [5,176].Criteria2Operator := -999, [5,176].Action := -999, [5,176].Label := -999, [5,176].Criteria1Value := -1000000.0, [5,176].Criteria2Value := -1000000.0, [5,176].ActionValue := -1000000.0, [5,177].Criteria1 := -999, [5,177].Criteria1Operator := -999, [5,177].Boolean := -999, [5,177].Criteria2 := -999, [5,177].Criteria2Operator := -999, [5,177].Action := -999, [5,177].Label := -999, [5,177].Criteria1Value := -1000000.0, [5,177].Criteria2Value := -1000000.0, [5,177].ActionValue := -1000000.0, [5,178].Criteria1 := -999, [5,178].Criteria1Operator := -999, [5,178].Boolean := -999, [5,178].Criteria2 := -999, [5,178].Criteria2Operator := -999, [5,178].Action := -999, [5,178].Label := -999, [5,178].Criteria1Value := -1000000.0, [5,178].Criteria2Value := -1000000.0, [5,178].ActionValue := -1000000.0, [5,179].Criteria1 := -999, [5,179].Criteria1Operator := -999, [5,179].Boolean := -999, [5,179].Criteria2 := -999, [5,179].Criteria2Operator := -999,
        [5,179].Action := -999, [5,179].Label := -999, [5,179].Criteria1Value := -1000000.0, [5,179].Criteria2Value := -1000000.0, [5,179].ActionValue := -1000000.0, [5,180].Criteria1 := -999, [5,180].Criteria1Operator := -999, [5,180].Boolean := -999, [5,180].Criteria2 := -999, [5,180].Criteria2Operator := -999, [5,180].Action := -999, [5,180].Label := -999, [5,180].Criteria1Value := -1000000.0, [5,180].Criteria2Value := -1000000.0, [5,180].ActionValue := -1000000.0, [5,181].Criteria1 := -999, [5,181].Criteria1Operator := -999, [5,181].Boolean := -999, [5,181].Criteria2 := -999, [5,181].Criteria2Operator := -999, [5,181].Action := -999, [5,181].Label := -999, [5,181].Criteria1Value := -1000000.0, [5,181].Criteria2Value := -1000000.0, [5,181].ActionValue := -1000000.0, [5,182].Criteria1 := -999, [5,182].Criteria1Operator := -999, [5,182].Boolean := -999, [5,182].Criteria2 := -999, [5,182].Criteria2Operator := -999, [5,182].Action := -999, [5,182].Label := -999, [5,182].Criteria1Value := -1000000.0, [5,182].Criteria2Value := -1000000.0, [5,182].ActionValue := -1000000.0, [5,183].Criteria1 := -999, [5,183].Criteria1Operator := -999, [5,183].Boolean := -999, [5,183].Criteria2 := -999, [5,183].Criteria2Operator := -999, [5,183].Action := -999, [5,183].Label := -999, [5,183].Criteria1Value := -1000000.0, [5,183].Criteria2Value := -1000000.0, [5,183].ActionValue := -1000000.0, [5,184].Criteria1 := -999, [5,184].Criteria1Operator := -999, [5,184].Boolean := -999, [5,184].Criteria2 := -999, [5,184].Criteria2Operator := -999, [5,184].Action := -999, [5,184].Label := -999, [5,184].Criteria1Value := -1000000.0, [5,184].Criteria2Value := -1000000.0, [5,184].ActionValue := -1000000.0, [5,185].Criteria1 := -999, [5,185].Criteria1Operator := -999, [5,185].Boolean := -999, [5,185].Criteria2 := -999, [5,185].Criteria2Operator := -999,
        [5,185].Action := -999, [5,185].Label := -999, [5,185].Criteria1Value := -1000000.0, [5,185].Criteria2Value := -1000000.0, [5,185].ActionValue := -1000000.0, [5,186].Criteria1 := -999, [5,186].Criteria1Operator := -999, [5,186].Boolean := -999, [5,186].Criteria2 := -999, [5,186].Criteria2Operator := -999, [5,186].Action := -999, [5,186].Label := -999, [5,186].Criteria1Value := -1000000.0, [5,186].Criteria2Value := -1000000.0, [5,186].ActionValue := -1000000.0, [5,187].Criteria1 := -999, [5,187].Criteria1Operator := -999, [5,187].Boolean := -999, [5,187].Criteria2 := -999, [5,187].Criteria2Operator := -999, [5,187].Action := -999, [5,187].Label := -999, [5,187].Criteria1Value := -1000000.0, [5,187].Criteria2Value := -1000000.0, [5,187].ActionValue := -1000000.0, [5,188].Criteria1 := -999, [5,188].Criteria1Operator := -999, [5,188].Boolean := -999, [5,188].Criteria2 := -999, [5,188].Criteria2Operator := -999, [5,188].Action := -999, [5,188].Label := -999, [5,188].Criteria1Value := -1000000.0, [5,188].Criteria2Value := -1000000.0, [5,188].ActionValue := -1000000.0, [5,189].Criteria1 := -999, [5,189].Criteria1Operator := -999, [5,189].Boolean := -999, [5,189].Criteria2 := -999, [5,189].Criteria2Operator := -999, [5,189].Action := -999, [5,189].Label := -999, [5,189].Criteria1Value := -1000000.0, [5,189].Criteria2Value := -1000000.0, [5,189].ActionValue := -1000000.0, [5,190].Criteria1 := -999, [5,190].Criteria1Operator := -999, [5,190].Boolean := -999, [5,190].Criteria2 := -999, [5,190].Criteria2Operator := -999, [5,190].Action := -999, [5,190].Label := -999, [5,190].Criteria1Value := -1000000.0, [5,190].Criteria2Value := -1000000.0, [5,190].ActionValue := -1000000.0, [5,191].Criteria1 := -999, [5,191].Criteria1Operator := -999, [5,191].Boolean := -999, [5,191].Criteria2 := -999, [5,191].Criteria2Operator := -999,
        [5,191].Action := -999, [5,191].Label := -999, [5,191].Criteria1Value := -1000000.0, [5,191].Criteria2Value := -1000000.0, [5,191].ActionValue := -1000000.0, [5,192].Criteria1 := -999, [5,192].Criteria1Operator := -999, [5,192].Boolean := -999, [5,192].Criteria2 := -999, [5,192].Criteria2Operator := -999, [5,192].Action := -999, [5,192].Label := -999, [5,192].Criteria1Value := -1000000.0, [5,192].Criteria2Value := -1000000.0, [5,192].ActionValue := -1000000.0, [5,193].Criteria1 := -999, [5,193].Criteria1Operator := -999, [5,193].Boolean := -999, [5,193].Criteria2 := -999, [5,193].Criteria2Operator := -999, [5,193].Action := -999, [5,193].Label := -999, [5,193].Criteria1Value := -1000000.0, [5,193].Criteria2Value := -1000000.0, [5,193].ActionValue := -1000000.0, [5,194].Criteria1 := -999, [5,194].Criteria1Operator := -999, [5,194].Boolean := -999, [5,194].Criteria2 := -999, [5,194].Criteria2Operator := -999, [5,194].Action := -999, [5,194].Label := -999, [5,194].Criteria1Value := -1000000.0, [5,194].Criteria2Value := -1000000.0, [5,194].ActionValue := -1000000.0, [5,195].Criteria1 := -999, [5,195].Criteria1Operator := -999, [5,195].Boolean := -999, [5,195].Criteria2 := -999, [5,195].Criteria2Operator := -999, [5,195].Action := -999, [5,195].Label := -999, [5,195].Criteria1Value := -1000000.0, [5,195].Criteria2Value := -1000000.0, [5,195].ActionValue := -1000000.0, [5,196].Criteria1 := -999, [5,196].Criteria1Operator := -999, [5,196].Boolean := -999, [5,196].Criteria2 := -999, [5,196].Criteria2Operator := -999, [5,196].Action := -999, [5,196].Label := -999, [5,196].Criteria1Value := -1000000.0, [5,196].Criteria2Value := -1000000.0, [5,196].ActionValue := -1000000.0, [5,197].Criteria1 := -999, [5,197].Criteria1Operator := -999, [5,197].Boolean := -999, [5,197].Criteria2 := -999, [5,197].Criteria2Operator := -999,
        [5,197].Action := -999, [5,197].Label := -999, [5,197].Criteria1Value := -1000000.0, [5,197].Criteria2Value := -1000000.0, [5,197].ActionValue := -1000000.0, [5,198].Criteria1 := -999, [5,198].Criteria1Operator := -999, [5,198].Boolean := -999, [5,198].Criteria2 := -999, [5,198].Criteria2Operator := -999, [5,198].Action := -999, [5,198].Label := -999, [5,198].Criteria1Value := -1000000.0, [5,198].Criteria2Value := -1000000.0, [5,198].ActionValue := -1000000.0, [5,199].Criteria1 := -999, [5,199].Criteria1Operator := -999, [5,199].Boolean := -999, [5,199].Criteria2 := -999, [5,199].Criteria2Operator := -999, [5,199].Action := -999, [5,199].Label := -999, [5,199].Criteria1Value := -1000000.0, [5,199].Criteria2Value := -1000000.0, [5,199].ActionValue := -1000000.0, [5,200].Criteria1 := -999, [5,200].Criteria1Operator := -999, [5,200].Boolean := -999, [5,200].Criteria2 := -999, [5,200].Criteria2Operator := -999, [5,200].Action := -999, [5,200].Label := -999, [5,200].Criteria1Value := -1000000.0, [5,200].Criteria2Value := -1000000.0, [5,200].ActionValue := -1000000.0, [5,201].Criteria1 := -999, [5,201].Criteria1Operator := -999, [5,201].Boolean := -999, [5,201].Criteria2 := -999, [5,201].Criteria2Operator := -999, [5,201].Action := -999, [5,201].Label := -999, [5,201].Criteria1Value := -1000000.0, [5,201].Criteria2Value := -1000000.0, [5,201].ActionValue := -1000000.0, [5,202].Criteria1 := -999, [5,202].Criteria1Operator := -999, [5,202].Boolean := -999, [5,202].Criteria2 := -999, [5,202].Criteria2Operator := -999, [5,202].Action := -999, [5,202].Label := -999, [5,202].Criteria1Value := -1000000.0, [5,202].Criteria2Value := -1000000.0, [5,202].ActionValue := -1000000.0, [5,203].Criteria1 := -999, [5,203].Criteria1Operator := -999, [5,203].Boolean := -999, [5,203].Criteria2 := -999, [5,203].Criteria2Operator := -999,
        [5,203].Action := -999, [5,203].Label := -999, [5,203].Criteria1Value := -1000000.0, [5,203].Criteria2Value := -1000000.0, [5,203].ActionValue := -1000000.0, [5,204].Criteria1 := -999, [5,204].Criteria1Operator := -999, [5,204].Boolean := -999, [5,204].Criteria2 := -999, [5,204].Criteria2Operator := -999, [5,204].Action := -999, [5,204].Label := -999, [5,204].Criteria1Value := -1000000.0, [5,204].Criteria2Value := -1000000.0, [5,204].ActionValue := -1000000.0, [5,205].Criteria1 := -999, [5,205].Criteria1Operator := -999, [5,205].Boolean := -999, [5,205].Criteria2 := -999, [5,205].Criteria2Operator := -999, [5,205].Action := -999, [5,205].Label := -999, [5,205].Criteria1Value := -1000000.0, [5,205].Criteria2Value := -1000000.0, [5,205].ActionValue := -1000000.0, [5,206].Criteria1 := -999, [5,206].Criteria1Operator := -999, [5,206].Boolean := -999, [5,206].Criteria2 := -999, [5,206].Criteria2Operator := -999, [5,206].Action := -999, [5,206].Label := -999, [5,206].Criteria1Value := -1000000.0, [5,206].Criteria2Value := -1000000.0, [5,206].ActionValue := -1000000.0, [5,207].Criteria1 := -999, [5,207].Criteria1Operator := -999, [5,207].Boolean := -999, [5,207].Criteria2 := -999, [5,207].Criteria2Operator := -999, [5,207].Action := -999, [5,207].Label := -999, [5,207].Criteria1Value := -1000000.0, [5,207].Criteria2Value := -1000000.0, [5,207].ActionValue := -1000000.0, [5,208].Criteria1 := -999, [5,208].Criteria1Operator := -999, [5,208].Boolean := -999, [5,208].Criteria2 := -999, [5,208].Criteria2Operator := -999, [5,208].Action := -999, [5,208].Label := -999, [5,208].Criteria1Value := -1000000.0, [5,208].Criteria2Value := -1000000.0, [5,208].ActionValue := -1000000.0, [5,209].Criteria1 := -999, [5,209].Criteria1Operator := -999, [5,209].Boolean := -999, [5,209].Criteria2 := -999, [5,209].Criteria2Operator := -999,
        [5,209].Action := -999, [5,209].Label := -999, [5,209].Criteria1Value := -1000000.0, [5,209].Criteria2Value := -1000000.0, [5,209].ActionValue := -1000000.0, [5,210].Criteria1 := -999, [5,210].Criteria1Operator := -999, [5,210].Boolean := -999, [5,210].Criteria2 := -999, [5,210].Criteria2Operator := -999, [5,210].Action := -999, [5,210].Label := -999, [5,210].Criteria1Value := -1000000.0, [5,210].Criteria2Value := -1000000.0, [5,210].ActionValue := -1000000.0, [5,211].Criteria1 := -999, [5,211].Criteria1Operator := -999, [5,211].Boolean := -999, [5,211].Criteria2 := -999, [5,211].Criteria2Operator := -999, [5,211].Action := -999, [5,211].Label := -999, [5,211].Criteria1Value := -1000000.0, [5,211].Criteria2Value := -1000000.0, [5,211].ActionValue := -1000000.0, [5,212].Criteria1 := -999, [5,212].Criteria1Operator := -999, [5,212].Boolean := -999, [5,212].Criteria2 := -999, [5,212].Criteria2Operator := -999, [5,212].Action := -999, [5,212].Label := -999, [5,212].Criteria1Value := -1000000.0, [5,212].Criteria2Value := -1000000.0, [5,212].ActionValue := -1000000.0, [5,213].Criteria1 := -999, [5,213].Criteria1Operator := -999, [5,213].Boolean := -999, [5,213].Criteria2 := -999, [5,213].Criteria2Operator := -999, [5,213].Action := -999, [5,213].Label := -999, [5,213].Criteria1Value := -1000000.0, [5,213].Criteria2Value := -1000000.0, [5,213].ActionValue := -1000000.0, [5,214].Criteria1 := -999, [5,214].Criteria1Operator := -999, [5,214].Boolean := -999, [5,214].Criteria2 := -999, [5,214].Criteria2Operator := -999, [5,214].Action := -999, [5,214].Label := -999, [5,214].Criteria1Value := -1000000.0, [5,214].Criteria2Value := -1000000.0, [5,214].ActionValue := -1000000.0, [5,215].Criteria1 := -999, [5,215].Criteria1Operator := -999, [5,215].Boolean := -999, [5,215].Criteria2 := -999, [5,215].Criteria2Operator := -999,
        [5,215].Action := -999, [5,215].Label := -999, [5,215].Criteria1Value := -1000000.0, [5,215].Criteria2Value := -1000000.0, [5,215].ActionValue := -1000000.0, [5,216].Criteria1 := -999, [5,216].Criteria1Operator := -999, [5,216].Boolean := -999, [5,216].Criteria2 := -999, [5,216].Criteria2Operator := -999, [5,216].Action := -999, [5,216].Label := -999, [5,216].Criteria1Value := -1000000.0, [5,216].Criteria2Value := -1000000.0, [5,216].ActionValue := -1000000.0, [5,217].Criteria1 := -999, [5,217].Criteria1Operator := -999, [5,217].Boolean := -999, [5,217].Criteria2 := -999, [5,217].Criteria2Operator := -999, [5,217].Action := -999, [5,217].Label := -999, [5,217].Criteria1Value := -1000000.0, [5,217].Criteria2Value := -1000000.0, [5,217].ActionValue := -1000000.0, [5,218].Criteria1 := -999, [5,218].Criteria1Operator := -999, [5,218].Boolean := -999, [5,218].Criteria2 := -999, [5,218].Criteria2Operator := -999, [5,218].Action := -999, [5,218].Label := -999, [5,218].Criteria1Value := -1000000.0, [5,218].Criteria2Value := -1000000.0, [5,218].ActionValue := -1000000.0, [5,219].Criteria1 := -999, [5,219].Criteria1Operator := -999, [5,219].Boolean := -999, [5,219].Criteria2 := -999, [5,219].Criteria2Operator := -999, [5,219].Action := -999, [5,219].Label := -999, [5,219].Criteria1Value := -1000000.0, [5,219].Criteria2Value := -1000000.0, [5,219].ActionValue := -1000000.0, [5,220].Criteria1 := -999, [5,220].Criteria1Operator := -999, [5,220].Boolean := -999, [5,220].Criteria2 := -999, [5,220].Criteria2Operator := -999, [5,220].Action := -999, [5,220].Label := -999, [5,220].Criteria1Value := -1000000.0, [5,220].Criteria2Value := -1000000.0, [5,220].ActionValue := -1000000.0, [5,221].Criteria1 := -999, [5,221].Criteria1Operator := -999, [5,221].Boolean := -999, [5,221].Criteria2 := -999, [5,221].Criteria2Operator := -999,
        [5,221].Action := -999, [5,221].Label := -999, [5,221].Criteria1Value := -1000000.0, [5,221].Criteria2Value := -1000000.0, [5,221].ActionValue := -1000000.0, [5,222].Criteria1 := -999, [5,222].Criteria1Operator := -999, [5,222].Boolean := -999, [5,222].Criteria2 := -999, [5,222].Criteria2Operator := -999, [5,222].Action := -999, [5,222].Label := -999, [5,222].Criteria1Value := -1000000.0, [5,222].Criteria2Value := -1000000.0, [5,222].ActionValue := -1000000.0, [5,223].Criteria1 := -999, [5,223].Criteria1Operator := -999, [5,223].Boolean := -999, [5,223].Criteria2 := -999, [5,223].Criteria2Operator := -999, [5,223].Action := -999, [5,223].Label := -999, [5,223].Criteria1Value := -1000000.0, [5,223].Criteria2Value := -1000000.0, [5,223].ActionValue := -1000000.0, [5,224].Criteria1 := -999, [5,224].Criteria1Operator := -999, [5,224].Boolean := -999, [5,224].Criteria2 := -999, [5,224].Criteria2Operator := -999, [5,224].Action := -999, [5,224].Label := -999, [5,224].Criteria1Value := -1000000.0, [5,224].Criteria2Value := -1000000.0, [5,224].ActionValue := -1000000.0, [5,225].Criteria1 := -999, [5,225].Criteria1Operator := -999, [5,225].Boolean := -999, [5,225].Criteria2 := -999, [5,225].Criteria2Operator := -999, [5,225].Action := -999, [5,225].Label := -999, [5,225].Criteria1Value := -1000000.0, [5,225].Criteria2Value := -1000000.0, [5,225].ActionValue := -1000000.0, [5,226].Criteria1 := -999, [5,226].Criteria1Operator := -999, [5,226].Boolean := -999, [5,226].Criteria2 := -999, [5,226].Criteria2Operator := -999, [5,226].Action := -999, [5,226].Label := -999, [5,226].Criteria1Value := -1000000.0, [5,226].Criteria2Value := -1000000.0, [5,226].ActionValue := -1000000.0, [5,227].Criteria1 := -999, [5,227].Criteria1Operator := -999, [5,227].Boolean := -999, [5,227].Criteria2 := -999, [5,227].Criteria2Operator := -999,
        [5,227].Action := -999, [5,227].Label := -999, [5,227].Criteria1Value := -1000000.0, [5,227].Criteria2Value := -1000000.0, [5,227].ActionValue := -1000000.0, [5,228].Criteria1 := -999, [5,228].Criteria1Operator := -999, [5,228].Boolean := -999, [5,228].Criteria2 := -999, [5,228].Criteria2Operator := -999, [5,228].Action := -999, [5,228].Label := -999, [5,228].Criteria1Value := -1000000.0, [5,228].Criteria2Value := -1000000.0, [5,228].ActionValue := -1000000.0, [5,229].Criteria1 := -999, [5,229].Criteria1Operator := -999, [5,229].Boolean := -999, [5,229].Criteria2 := -999, [5,229].Criteria2Operator := -999, [5,229].Action := -999, [5,229].Label := -999, [5,229].Criteria1Value := -1000000.0, [5,229].Criteria2Value := -1000000.0, [5,229].ActionValue := -1000000.0, [5,230].Criteria1 := -999, [5,230].Criteria1Operator := -999, [5,230].Boolean := -999, [5,230].Criteria2 := -999, [5,230].Criteria2Operator := -999, [5,230].Action := -999, [5,230].Label := -999, [5,230].Criteria1Value := -1000000.0, [5,230].Criteria2Value := -1000000.0, [5,230].ActionValue := -1000000.0, [5,231].Criteria1 := -999, [5,231].Criteria1Operator := -999, [5,231].Boolean := -999, [5,231].Criteria2 := -999, [5,231].Criteria2Operator := -999, [5,231].Action := -999, [5,231].Label := -999, [5,231].Criteria1Value := -1000000.0, [5,231].Criteria2Value := -1000000.0, [5,231].ActionValue := -1000000.0, [5,232].Criteria1 := -999, [5,232].Criteria1Operator := -999, [5,232].Boolean := -999, [5,232].Criteria2 := -999, [5,232].Criteria2Operator := -999, [5,232].Action := -999, [5,232].Label := -999, [5,232].Criteria1Value := -1000000.0, [5,232].Criteria2Value := -1000000.0, [5,232].ActionValue := -1000000.0, [5,233].Criteria1 := -999, [5,233].Criteria1Operator := -999, [5,233].Boolean := -999, [5,233].Criteria2 := -999, [5,233].Criteria2Operator := -999,
        [5,233].Action := -999, [5,233].Label := -999, [5,233].Criteria1Value := -1000000.0, [5,233].Criteria2Value := -1000000.0, [5,233].ActionValue := -1000000.0, [5,234].Criteria1 := -999, [5,234].Criteria1Operator := -999, [5,234].Boolean := -999, [5,234].Criteria2 := -999, [5,234].Criteria2Operator := -999, [5,234].Action := -999, [5,234].Label := -999, [5,234].Criteria1Value := -1000000.0, [5,234].Criteria2Value := -1000000.0, [5,234].ActionValue := -1000000.0, [5,235].Criteria1 := -999, [5,235].Criteria1Operator := -999, [5,235].Boolean := -999, [5,235].Criteria2 := -999, [5,235].Criteria2Operator := -999, [5,235].Action := -999, [5,235].Label := -999, [5,235].Criteria1Value := -1000000.0, [5,235].Criteria2Value := -1000000.0, [5,235].ActionValue := -1000000.0, [5,236].Criteria1 := -999, [5,236].Criteria1Operator := -999, [5,236].Boolean := -999, [5,236].Criteria2 := -999, [5,236].Criteria2Operator := -999, [5,236].Action := -999, [5,236].Label := -999, [5,236].Criteria1Value := -1000000.0, [5,236].Criteria2Value := -1000000.0, [5,236].ActionValue := -1000000.0, [5,237].Criteria1 := -999, [5,237].Criteria1Operator := -999, [5,237].Boolean := -999, [5,237].Criteria2 := -999, [5,237].Criteria2Operator := -999, [5,237].Action := -999, [5,237].Label := -999, [5,237].Criteria1Value := -1000000.0, [5,237].Criteria2Value := -1000000.0, [5,237].ActionValue := -1000000.0, [5,238].Criteria1 := -999, [5,238].Criteria1Operator := -999, [5,238].Boolean := -999, [5,238].Criteria2 := -999, [5,238].Criteria2Operator := -999, [5,238].Action := -999, [5,238].Label := -999, [5,238].Criteria1Value := -1000000.0, [5,238].Criteria2Value := -1000000.0, [5,238].ActionValue := -1000000.0, [5,239].Criteria1 := -999, [5,239].Criteria1Operator := -999, [5,239].Boolean := -999, [5,239].Criteria2 := -999, [5,239].Criteria2Operator := -999,
        [5,239].Action := -999, [5,239].Label := -999, [5,239].Criteria1Value := -1000000.0, [5,239].Criteria2Value := -1000000.0, [5,239].ActionValue := -1000000.0, [5,240].Criteria1 := -999, [5,240].Criteria1Operator := -999, [5,240].Boolean := -999, [5,240].Criteria2 := -999, [5,240].Criteria2Operator := -999, [5,240].Action := -999, [5,240].Label := -999, [5,240].Criteria1Value := -1000000.0, [5,240].Criteria2Value := -1000000.0, [5,240].ActionValue := -1000000.0, [5,241].Criteria1 := -999, [5,241].Criteria1Operator := -999, [5,241].Boolean := -999, [5,241].Criteria2 := -999, [5,241].Criteria2Operator := -999, [5,241].Action := -999, [5,241].Label := -999, [5,241].Criteria1Value := -1000000.0, [5,241].Criteria2Value := -1000000.0, [5,241].ActionValue := -1000000.0, [5,242].Criteria1 := -999, [5,242].Criteria1Operator := -999, [5,242].Boolean := -999, [5,242].Criteria2 := -999, [5,242].Criteria2Operator := -999, [5,242].Action := -999, [5,242].Label := -999, [5,242].Criteria1Value := -1000000.0, [5,242].Criteria2Value := -1000000.0, [5,242].ActionValue := -1000000.0, [5,243].Criteria1 := -999, [5,243].Criteria1Operator := -999, [5,243].Boolean := -999, [5,243].Criteria2 := -999, [5,243].Criteria2Operator := -999, [5,243].Action := -999, [5,243].Label := -999, [5,243].Criteria1Value := -1000000.0, [5,243].Criteria2Value := -1000000.0, [5,243].ActionValue := -1000000.0, [5,244].Criteria1 := -999, [5,244].Criteria1Operator := -999, [5,244].Boolean := -999, [5,244].Criteria2 := -999, [5,244].Criteria2Operator := -999, [5,244].Action := -999, [5,244].Label := -999, [5,244].Criteria1Value := -1000000.0, [5,244].Criteria2Value := -1000000.0, [5,244].ActionValue := -1000000.0, [5,245].Criteria1 := -999, [5,245].Criteria1Operator := -999, [5,245].Boolean := -999, [5,245].Criteria2 := -999, [5,245].Criteria2Operator := -999,
        [5,245].Action := -999, [5,245].Label := -999, [5,245].Criteria1Value := -1000000.0, [5,245].Criteria2Value := -1000000.0, [5,245].ActionValue := -1000000.0, [5,246].Criteria1 := -999, [5,246].Criteria1Operator := -999, [5,246].Boolean := -999, [5,246].Criteria2 := -999, [5,246].Criteria2Operator := -999, [5,246].Action := -999, [5,246].Label := -999, [5,246].Criteria1Value := -1000000.0, [5,246].Criteria2Value := -1000000.0, [5,246].ActionValue := -1000000.0, [5,247].Criteria1 := -999, [5,247].Criteria1Operator := -999, [5,247].Boolean := -999, [5,247].Criteria2 := -999, [5,247].Criteria2Operator := -999, [5,247].Action := -999, [5,247].Label := -999, [5,247].Criteria1Value := -1000000.0, [5,247].Criteria2Value := -1000000.0, [5,247].ActionValue := -1000000.0, [5,248].Criteria1 := -999, [5,248].Criteria1Operator := -999, [5,248].Boolean := -999, [5,248].Criteria2 := -999, [5,248].Criteria2Operator := -999, [5,248].Action := -999, [5,248].Label := -999, [5,248].Criteria1Value := -1000000.0, [5,248].Criteria2Value := -1000000.0, [5,248].ActionValue := -1000000.0, [5,249].Criteria1 := -999, [5,249].Criteria1Operator := -999, [5,249].Boolean := -999, [5,249].Criteria2 := -999, [5,249].Criteria2Operator := -999, [5,249].Action := -999, [5,249].Label := -999, [5,249].Criteria1Value := -1000000.0, [5,249].Criteria2Value := -1000000.0, [5,249].ActionValue := -1000000.0, [5,250].Criteria1 := -999, [5,250].Criteria1Operator := -999, [5,250].Boolean := -999, [5,250].Criteria2 := -999, [5,250].Criteria2Operator := -999, [5,250].Action := -999, [5,250].Label := -999, [5,250].Criteria1Value := -1000000.0, [5,250].Criteria2Value := -1000000.0, [5,250].ActionValue := -1000000.0);   // Operation Table
        [0,0]   // Null Step
        [1,0]   // Null Step
        [2,0]   // Null Step
        [3,0]   // Null Step
        [4,0]   // Null Step
        [5,0]   // Null Step
   Options : Options := (WI102 := 1, AI101_AI102_AI103 := 1, Tank250 := 1, CCP_Report := 1, TF3S := 1);   // Options List
   PCDateTime : DINT[7] := ([0] := 2026, [1] := 7, [2] := 24, [3] := 11, [4] := 30, [5] := 6, [6] := -1);   // Date/Time Array from PC
   PcToPLCHeartBeat : BOOL;   // PC to PLC communication heartbeat Set to 1 by HMI Reset to 0 by plc
   PCV001 : ALIAS FOR AnalogPoint[3];   // Retentate Pressure Control Valve Position
   PCV001_AO : ALIAS FOR AnalogOutput[0];   // Retentate Pressure Control Valve Setpoint
   PCV001_Calib : PCV_Calib;   // PCV001 Position Calibration
   PCV001_Control : PCV_Control := (FullOpenResetTimer.PRE := 1000, FullCloseSP := 100.0, FullCloseResetTimer.PRE := 1000, ClosedStatusSP := 95.0);   // PCV001 Control UDT
   PCV001_CVTune : CVTune := (ClosedRaw := 23479.0, OpenRaw := 17404.0, MaxOutput := 100.0, MinTimer.PRE := 5000, MaxTimer.PRE := 5000);
   PCV001_PID : PCV := (PV := -0.08230453, CV := 2.2879825, OpenRawValue := 17404.0, ClosedRawValue := 23479.0);   // PCV001 PID Management
   PCV001_SIG : ALIAS FOR DigitalPoint[102];
   PCV101 : ALIAS FOR AnalogPoint[4];   // Filtrate Pressure Control Valve Position
   PCV101_AO : ALIAS FOR AnalogOutput[1];   // FiltratePressure Control Valve Setpoint
   PCV101_Calib : PCV_Calib;   // PCV101 Position Calibration
   PCV101_Control : PCV_Control := (FullOpenSP := 100.0, FullOpenResetTimer.PRE := 1000, FullCloseResetTimer.PRE := 1000, ClosedStatusSP := 95.0);   // PCV101 Control UDT
   PCV101_CVTune : CVTune := (ClosedRaw := 17268.0, OpenRaw := 23352.0, MaxOutput := 100.0, MinTimer.PRE := 5000, MaxTimer.PRE := 5000);
   PCV101_PID : PCV := (PV := 99.52334, CV := 86.55756, OpenRawValue := 23352.0, ClosedRawValue := 17268.0);   // PCV101 PID Management
   PCV101_SIG : ALIAS FOR DigitalPoint[103];
   PERM : ALIAS FOR AnalogPoint[46];   // Membrane Permeability
   PERMAlarm : ALIAS FOR AlarmAnalog[46];   // PERM Alarm
   Phase : Phases[6] := ([0].JumpStep := 62, [0].StartStep := 1, [0].TotalSteps := 60, [0].ActualStep := 61, [1].Stop := 1, [1].JumpStep := 4, [1].StartStep := 1, [1].Crit1MetTime := 16, [1].TotalSteps := 10, [1].ActualStep := 3, [2].Stop := 1, [2].JumpStep := 6, [2].StartStep := 1, [2].ActualStep := 5, [3].Stop := 1, [3].JumpStep := 11, [3].StartStep := 1, [3].TotalSteps := 9, [3].ActualStep := 10, [4].JumpStep := 23, [4].StartStep := 1, [4].TotalSteps := 21, [4].ActualStep := 22, [5].JumpStep := 70, [5].StartStep := 1, [5].ActualStep := 69);   // Phase Control Array
   Phase0 : ALIAS FOR Phase[0];   // Phase 0
   Phase0_PauseTime : ALIAS FOR Timers[12];   // Phase 0 Pause Time
   Phase0_StepTime : ALIAS FOR Timers[6];   // Phase 0 Step Time
   Phase0_Totalizer_Feed : ALIAS FOR PhaseTotalizer[0];   // Phase 0 Total Feed
   Phase0_Totalizer_Filtrate : ALIAS FOR PhaseTotalizer[6];   // Phase 0 Total Filtrate
   Phase0_Totalizer_Retentate : ALIAS FOR PhaseTotalizer[12];   // Phase 0 Total Retentate
   Phase0_TotalTime : ALIAS FOR Timers[0];   // Phase 0 Total Time
   Phase1 : ALIAS FOR Phase[1];   // Phase 1
   Phase1_PauseTime : ALIAS FOR Timers[13];   // Phase 1 Pause Time
   Phase1_StepTime : ALIAS FOR Timers[7];   // Phase 1 Step Time
   Phase1_Totalizer_Feed : ALIAS FOR PhaseTotalizer[1];   // Phase 1 Total Feed
   Phase1_Totalizer_Filtrate : ALIAS FOR PhaseTotalizer[7];   // Phase 1 Total Filtrate
   Phase1_Totalizer_Retentate : ALIAS FOR PhaseTotalizer[13];   // Phase 1 Total Retentate
   Phase1_TotalTime : ALIAS FOR Timers[1];   // Phase 1 Total Time
   Phase2 : ALIAS FOR Phase[2];   // Phase 2
   Phase2_PauseTime : ALIAS FOR Timers[14];   // Phase 2 Pause Time
   Phase2_StepTime : ALIAS FOR Timers[8];   // Phase 2 Step Time
   Phase2_Totalizer_Feed : ALIAS FOR PhaseTotalizer[2];   // Phase 2 Total Feed
   Phase2_Totalizer_Filtrate : ALIAS FOR PhaseTotalizer[8];   // Phase 2 Total Filtrate
   Phase2_Totalizer_Retentate : ALIAS FOR PhaseTotalizer[14];   // Phase 2 Total Retentate
   Phase2_TotalTime : ALIAS FOR Timers[2];   // Phase 2 Total Time
   Phase3 : ALIAS FOR Phase[3];   // Phase 3
   Phase3_PauseTime : ALIAS FOR Timers[15];   // Phase 3 Pause Time
   Phase3_StepTime : ALIAS FOR Timers[9];   // Phase 3 Step Time
   Phase3_Totalizer_Feed : ALIAS FOR PhaseTotalizer[3];   // Phase 3 Total Feed
   Phase3_Totalizer_Filtrate : ALIAS FOR PhaseTotalizer[9];   // Phase 3 Total Filtrate
   Phase3_Totalizer_Retentate : ALIAS FOR PhaseTotalizer[15];   // Phase 3 Total Retentate
   Phase3_TotalTime : ALIAS FOR Timers[3];   // Phase 3 Total Time
   Phase4 : ALIAS FOR Phase[4];   // Phase 4
   Phase4_PauseTime : ALIAS FOR Timers[16];   // Phase 4 Pause Time
   Phase4_StepTime : ALIAS FOR Timers[10];   // Phase 4 Step Time
   Phase4_Totalizer_Feed : ALIAS FOR PhaseTotalizer[4];   // Phase 4 Total Feed
   Phase4_Totalizer_Filtrate : ALIAS FOR PhaseTotalizer[10];   // Phase 4 Total Filtrate
   Phase4_Totalizer_Retentate : ALIAS FOR PhaseTotalizer[16];   // Phase 4 Total Retentate
   Phase4_TotalTime : ALIAS FOR Timers[4];   // Phase 4 Total Time
   Phase5 : ALIAS FOR Phase[5];   // Phase 5
   Phase5_PauseTime : ALIAS FOR Timers[17];   // Phase 5 Pause Time
   Phase5_StepTime : ALIAS FOR Timers[11];   // Phase 5 Step Time
   Phase5_Totalizer_Feed : ALIAS FOR PhaseTotalizer[5];   // Phase 5 Total Feed
   Phase5_Totalizer_Filtrate : ALIAS FOR PhaseTotalizer[11];   // Phase 5 Total Filtrate
   Phase5_Totalizer_Retentate : ALIAS FOR PhaseTotalizer[17];   // Phase 5 Total Retentate
   Phase5_TotalTime : ALIAS FOR Timers[5];   // Phase 5 Total Time
   PhaseTotalizer : PhaseTotalizer[18] := ([0].Enable := 1, [0].PVscale := 60.0, [0].Title := 'Phase0 Vol', [0].EGU := 'L', [0].EnableCfg := 1, [0].SourceAddressCfg := 42, [1].Enable := 1, [1].PVscale := 60.0, [1].Title := 'Phase1 Vol', [1].EGU := 'L', [1].EnableCfg := 1, [1].SourceAddressCfg := 42, [2].PVscale := 60.0, [2].Title := 'Phase2 Vol', [2].EGU := 'L', [2].EnableCfg := 1, [2].SourceAddressCfg := 42, [3].PVscale := 60.0, [3].Title := 'Phase3 Vol', [3].EGU := 'L', [3].EnableCfg := 1, [3].SourceAddressCfg := 42, [4].PVscale := 60.0, [4].Title := 'Phase4 Vol', [4].EGU := 'L', [4].EnableCfg := 1, [4].SourceAddressCfg := 42, [5].PVscale := 60.0, [5].Title := 'Phase5 Vol', [5].EGU := 'L', [5].EnableCfg := 1, [5].SourceAddressCfg := 42, [6].Enable := 1, [6].PVscale := 60.0, [6].Title := 'Phase0 Vol', [6].EGU := 'L', [6].EnableCfg := 1, [6].SourceAddressCfg := 2, [7].PVscale := 60.0, [7].Title := 'Phase1 Vol', [7].EGU := 'L', [7].EnableCfg := 1, [7].SourceAddressCfg := 2, [8].PVscale := 60.0, [8].Title := 'Phase2 Vol', [8].EGU := 'L', [8].EnableCfg := 1, [8].SourceAddressCfg := 2, [9].PVscale := 60.0, [9].Title := 'Phase3 Vol', [9].EGU := 'L', [9].EnableCfg := 1, [9].SourceAddressCfg := 2, [10].PVscale := 60.0, [10].Title := 'Phase4 Vol', [10].EGU := 'L', [10].EnableCfg := 1, [10].SourceAddressCfg := 2, [11].PVscale := 60.0, [11].Title := 'Phase5 Vol',
        [11].EGU := 'L', [11].EnableCfg := 1, [11].SourceAddressCfg := 2, [12].StepReset := 1, [12].PVscale := 60.0, [12].SourceAddressCfg := 17, [13].StepReset := 1, [13].PVscale := 60.0, [13].SourceAddressCfg := 17, [14].StepReset := 1, [14].PVscale := 60.0, [14].SourceAddressCfg := 17, [15].StepReset := 1, [15].PVscale := 60.0, [15].SourceAddressCfg := 17, [16].StepReset := 1, [16].PVscale := 60.0, [16].SourceAddressCfg := 17, [17].StepReset := 1, [17].PVscale := 60.0, [17].SourceAddressCfg := 17);   // Phase Totalizers Array
        [10]   // Phase 4 Totalizer 2
        [11]   // Phase 5 Totalizer 2
        [0]   // Phase 0 Totalizer 1
        [1]   // Phase 1 Totalizer 1
        [2]   // Phase 2 Totalizer 1
        [3]   // Phase 3 Totalizer 1
        [4]   // Phase 4 Totalizer 1
        [5]   // Phase 5 Totalizer 1
        [6]   // Phase 0 Totalizer 2
        [7]   // Phase 1 Totalizer 2
        [8]   // Phase 2 Totalizer 2
        [9]   // Phase 3 Totalizer 2
   PhaseTotalizer_Storage : PhaseTotalizer[6,18] := ([0,0].Enable := 1, [0,0].PVscale := 60.0, [0,0].Title := 'Phase0 Vol', [0,0].EGU := 'L', [0,0].EnableCfg := 1, [0,0].SourceAddressCfg := 40, [0,1].Enable := 1, [0,1].PVscale := 60.0, [0,1].Title := 'Phase1 Vol', [0,1].EGU := 'L', [0,1].EnableCfg := 1, [0,1].SourceAddressCfg := 40, [0,2].PVscale := 60.0, [0,2].Title := 'Phase2 Vol', [0,2].EGU := 'L', [0,2].EnableCfg := 1, [0,2].SourceAddressCfg := 40, [0,3].PVscale := 60.0, [0,3].Title := 'Phase3 Vol', [0,3].EGU := 'L', [0,3].EnableCfg := 1, [0,3].SourceAddressCfg := 40, [0,4].PVscale := 60.0, [0,4].Title := 'Phase4 Vol', [0,4].EGU := 'L', [0,4].EnableCfg := 1, [0,4].SourceAddressCfg := 40, [0,5].PVscale := 60.0, [0,5].Title := 'Phase5 Vol', [0,5].EGU := 'L', [0,5].EnableCfg := 1, [0,5].SourceAddressCfg := 40, [0,6].Enable := 1, [0,6].PVscale := 60.0, [0,6].Title := 'Phase0 CVs', [0,6].EGU := 'CVs', [0,6].EnableCfg := 1, [0,6].SourceTypeCfg := 1, [0,7].PVscale := 60.0, [0,7].Title := 'Phase1 CVs', [0,7].EGU := 'CVs', [0,7].EnableCfg := 1, [0,7].SourceTypeCfg := 1, [0,8].PVscale := 60.0, [0,8].Title := 'Phase2 CVs', [0,8].EGU := 'CVs', [0,8].EnableCfg := 1, [0,8].SourceTypeCfg := 1, [0,9].PVscale := 60.0, [0,9].Title := 'Phase3 CVs', [0,9].EGU := 'CVs', [0,9].EnableCfg := 1, [0,9].SourceTypeCfg := 1, [0,10].PVscale := 60.0, [0,10].Title := 'Phase4 CVs', [0,10].EGU := 'CVs', [0,10].EnableCfg := 1, [0,10].SourceTypeCfg := 1, [0,11].PVscale := 60.0, [0,11].Title := 'Phase5 CVs',
        [0,11].EGU := 'CVs', [0,11].EnableCfg := 1, [0,11].SourceTypeCfg := 1, [1,0].Enable := 1, [1,0].Phase := 10.166667, [1,0].Step := 9.333332, [1,0].Procedure := 10.166667, [1,0].PVscale := 60.0, [1,0].Title := 'Phase0 Vol', [1,0].EGU := 'L', [1,0].EnableCfg := 1, [1,0].SourceAddressCfg := 42, [1,1].Enable := 1, [1,1].PVscale := 60.0, [1,1].Title := 'Phase1 Vol', [1,1].EGU := 'L', [1,1].EnableCfg := 1, [1,1].SourceAddressCfg := 42, [1,2].PVscale := 60.0, [1,2].Title := 'Phase2 Vol', [1,2].EGU := 'L', [1,2].EnableCfg := 1, [1,2].SourceAddressCfg := 42, [1,3].PVscale := 60.0, [1,3].Title := 'Phase3 Vol', [1,3].EGU := 'L', [1,3].EnableCfg := 1, [1,3].SourceAddressCfg := 42, [1,4].PVscale := 60.0, [1,4].Title := 'Phase4 Vol', [1,4].EGU := 'L', [1,4].EnableCfg := 1, [1,4].SourceAddressCfg := 42, [1,5].PVscale := 60.0, [1,5].Title := 'Phase5 Vol', [1,5].EGU := 'L', [1,5].EnableCfg := 1, [1,5].SourceAddressCfg := 42, [1,6].Enable := 1, [1,6].PV := 0.01201648, [1,6].PVscale := 60.0, [1,6].PVsec := 0.00020027466, [1,6].Title := 'Phase0 Vol', [1,6].EGU := 'L', [1,6].EnableCfg := 1, [1,6].SourceAddressCfg := 2, [1,7].PV := 0.01201648, [1,7].PVscale := 60.0, [1,7].PVsec := 0.00020027466, [1,7].Title := 'Phase1 Vol', [1,7].EGU := 'L', [1,7].EnableCfg := 1, [1,7].SourceAddressCfg := 2, [1,8].PV := 0.01201648, [1,8].PVscale := 60.0, [1,8].PVsec := 0.00020027466, [1,8].Title := 'Phase2 Vol', [1,8].EGU := 'L', [1,8].EnableCfg := 1, [1,8].SourceAddressCfg := 2,
        [1,9].PV := 0.01201648, [1,9].PVscale := 60.0, [1,9].PVsec := 0.00020027466, [1,9].Title := 'Phase3 Vol', [1,9].EGU := 'L', [1,9].EnableCfg := 1, [1,9].SourceAddressCfg := 2, [1,10].PV := 0.01201648, [1,10].PVscale := 60.0, [1,10].PVsec := 0.00020027466, [1,10].Title := 'Phase4 Vol', [1,10].EGU := 'L', [1,10].EnableCfg := 1, [1,10].SourceAddressCfg := 2, [1,11].PV := 0.01201648, [1,11].PVscale := 60.0, [1,11].PVsec := 0.00020027466, [1,11].Title := 'Phase5 Vol', [1,11].EGU := 'L', [1,11].EnableCfg := 1, [1,11].SourceAddressCfg := 2, [1,12].PVscale := 60.0, [1,12].SourceAddressCfg := 17, [1,13].PVscale := 60.0, [1,13].SourceAddressCfg := 17, [1,14].PVscale := 60.0, [1,14].SourceAddressCfg := 17, [1,15].PVscale := 60.0, [1,15].SourceAddressCfg := 17, [1,16].PVscale := 60.0, [1,16].SourceAddressCfg := 17, [1,17].PVscale := 60.0, [1,17].SourceAddressCfg := 17, [2,0].Enable := 1, [2,0].PVscale := 60.0, [2,0].Title := 'Phase0 Vol', [2,0].EGU := 'L', [2,0].EnableCfg := 1, [2,0].SourceAddressCfg := 42, [2,1].Enable := 1, [2,1].PVscale := 60.0, [2,1].Title := 'Phase1 Vol', [2,1].EGU := 'L', [2,1].EnableCfg := 1, [2,1].SourceAddressCfg := 42, [2,2].PVscale := 60.0, [2,2].Title := 'Phase2 Vol', [2,2].EGU := 'L', [2,2].EnableCfg := 1, [2,2].SourceAddressCfg := 42, [2,3].PVscale := 60.0, [2,3].Title := 'Phase3 Vol', [2,3].EGU := 'L', [2,3].EnableCfg := 1, [2,3].SourceAddressCfg := 42, [2,4].PVscale := 60.0, [2,4].Title := 'Phase4 Vol', [2,4].EGU := 'L', [2,4].EnableCfg := 1, [2,4].SourceAddressCfg := 42,
        [2,5].PVscale := 60.0, [2,5].Title := 'Phase5 Vol', [2,5].EGU := 'L', [2,5].EnableCfg := 1, [2,5].SourceAddressCfg := 42, [2,6].Enable := 1, [2,6].PV := -6.249523, [2,6].PVscale := 60.0, [2,6].Title := 'Phase0 Vol', [2,6].EGU := 'L', [2,6].EnableCfg := 1, [2,6].SourceAddressCfg := 2, [2,7].PV := -6.249523, [2,7].PVscale := 60.0, [2,7].Title := 'Phase1 Vol', [2,7].EGU := 'L', [2,7].EnableCfg := 1, [2,7].SourceAddressCfg := 2, [2,8].PV := -6.249523, [2,8].PVscale := 60.0, [2,8].Title := 'Phase2 Vol', [2,8].EGU := 'L', [2,8].EnableCfg := 1, [2,8].SourceAddressCfg := 2, [2,9].PV := -6.249523, [2,9].PVscale := 60.0, [2,9].Title := 'Phase3 Vol', [2,9].EGU := 'L', [2,9].EnableCfg := 1, [2,9].SourceAddressCfg := 2, [2,10].PV := -6.249523, [2,10].PVscale := 60.0, [2,10].Title := 'Phase4 Vol', [2,10].EGU := 'L', [2,10].EnableCfg := 1, [2,10].SourceAddressCfg := 2, [2,11].PV := -6.249523, [2,11].PVscale := 60.0, [2,11].Title := 'Phase5 Vol', [2,11].EGU := 'L', [2,11].EnableCfg := 1, [2,11].SourceAddressCfg := 2, [3,0].PV := 48.590927, [3,0].PVscale := 60.0, [3,0].PVsec := 0.8098488, [3,0].EnableCfg := 1, [3,0].SourceAddressCfg := 40, [3,1].PV := 48.590927, [3,1].PVscale := 60.0, [3,1].PVsec := 0.8098488, [3,1].EnableCfg := 1, [3,1].SourceAddressCfg := 40, [3,2].PV := 48.590927, [3,2].PVscale := 60.0, [3,2].PVsec := 0.8098488, [3,2].EnableCfg := 1, [3,2].SourceAddressCfg := 40, [3,3].PV := 48.590927, [3,3].PVscale := 60.0, [3,3].PVsec := 0.8098488,
        [3,3].EnableCfg := 1, [3,3].SourceAddressCfg := 40, [3,4].PV := 48.590927, [3,4].PVscale := 60.0, [3,4].PVsec := 0.8098488, [3,4].EnableCfg := 1, [3,4].SourceAddressCfg := 40, [3,5].PV := 48.590927, [3,5].PVscale := 60.0, [3,5].PVsec := 0.8098488, [3,5].EnableCfg := 1, [3,5].SourceAddressCfg := 40, [3,6].PV := 4.8590927, [3,6].PVscale := 60.0, [3,6].PVsec := 0.080984876, [3,6].EnableCfg := 1, [3,6].SourceTypeCfg := 1, [3,7].PV := 4.8590927, [3,7].PVscale := 60.0, [3,7].PVsec := 0.080984876, [3,7].EnableCfg := 1, [3,7].SourceTypeCfg := 1, [3,8].PV := 4.8590927, [3,8].PVscale := 60.0, [3,8].PVsec := 0.080984876, [3,8].EnableCfg := 1, [3,8].SourceTypeCfg := 1, [3,9].PV := 4.8590927, [3,9].PVscale := 60.0, [3,9].PVsec := 0.080984876, [3,9].EnableCfg := 1, [3,9].SourceTypeCfg := 1, [3,10].PV := 4.8590927, [3,10].PVscale := 60.0, [3,10].PVsec := 0.080984876, [3,10].EnableCfg := 1, [3,10].SourceTypeCfg := 1, [3,11].PV := 4.8590927, [3,11].PVscale := 60.0, [3,11].PVsec := 0.080984876, [3,11].EnableCfg := 1, [3,11].SourceTypeCfg := 1, [4,0].Enable := 1, [4,0].PVscale := 60.0, [4,0].Title := 'Phase0 Vol', [4,0].EGU := 'L', [4,0].EnableCfg := 1, [4,0].SourceAddressCfg := 40, [4,1].Enable := 1, [4,1].PVscale := 60.0, [4,1].Title := 'Phase1 Vol', [4,1].EGU := 'L', [4,1].EnableCfg := 1, [4,1].SourceAddressCfg := 40, [4,2].PVscale := 60.0, [4,2].Title := 'Phase2 Vol', [4,2].EGU := 'L', [4,2].EnableCfg := 1, [4,2].SourceAddressCfg := 40, [4,3].PVscale := 60.0,
        [4,3].Title := 'Phase3 Vol', [4,3].EGU := 'L', [4,3].EnableCfg := 1, [4,3].SourceAddressCfg := 40, [4,4].PVscale := 60.0, [4,4].Title := 'Phase4 Vol', [4,4].EGU := 'L', [4,4].EnableCfg := 1, [4,4].SourceAddressCfg := 40, [4,5].PVscale := 60.0, [4,5].Title := 'Phase5 Vol', [4,5].EGU := 'L', [4,5].EnableCfg := 1, [4,5].SourceAddressCfg := 40, [4,6].Enable := 1, [4,6].PVscale := 60.0, [4,6].Title := 'Phase0 CVs', [4,6].EGU := 'CVs', [4,6].EnableCfg := 1, [4,6].SourceTypeCfg := 1, [4,7].PVscale := 60.0, [4,7].Title := 'Phase1 CVs', [4,7].EGU := 'CVs', [4,7].EnableCfg := 1, [4,7].SourceTypeCfg := 1, [4,8].PVscale := 60.0, [4,8].Title := 'Phase2 CVs', [4,8].EGU := 'CVs', [4,8].EnableCfg := 1, [4,8].SourceTypeCfg := 1, [4,9].PVscale := 60.0, [4,9].Title := 'Phase3 CVs', [4,9].EGU := 'CVs', [4,9].EnableCfg := 1, [4,9].SourceTypeCfg := 1, [4,10].PVscale := 60.0, [4,10].Title := 'Phase4 CVs', [4,10].EGU := 'CVs', [4,10].EnableCfg := 1, [4,10].SourceTypeCfg := 1, [4,11].PVscale := 60.0, [4,11].Title := 'Phase5 CVs', [4,11].EGU := 'CVs', [4,11].EnableCfg := 1, [4,11].SourceTypeCfg := 1, [5,0].Enable := 1, [5,0].PVscale := 60.0, [5,0].Title := 'Phase0 Vol', [5,0].EGU := 'L', [5,0].EnableCfg := 1, [5,0].SourceAddressCfg := 40, [5,1].Enable := 1, [5,1].PVscale := 60.0, [5,1].Title := 'Phase1 Vol', [5,1].EGU := 'L', [5,1].EnableCfg := 1, [5,1].SourceAddressCfg := 40, [5,2].PVscale := 60.0, [5,2].Title := 'Phase2 Vol', [5,2].EGU := 'L',
        [5,2].EnableCfg := 1, [5,2].SourceAddressCfg := 40, [5,3].PVscale := 60.0, [5,3].Title := 'Phase3 Vol', [5,3].EGU := 'L', [5,3].EnableCfg := 1, [5,3].SourceAddressCfg := 40, [5,4].PVscale := 60.0, [5,4].Title := 'Phase4 Vol', [5,4].EGU := 'L', [5,4].EnableCfg := 1, [5,4].SourceAddressCfg := 40, [5,5].PVscale := 60.0, [5,5].Title := 'Phase5 Vol', [5,5].EGU := 'L', [5,5].EnableCfg := 1, [5,5].SourceAddressCfg := 40, [5,6].Enable := 1, [5,6].PVscale := 60.0, [5,6].Title := 'Phase0 CVs', [5,6].EGU := 'CVs', [5,6].EnableCfg := 1, [5,6].SourceTypeCfg := 1, [5,7].PVscale := 60.0, [5,7].Title := 'Phase1 CVs', [5,7].EGU := 'CVs', [5,7].EnableCfg := 1, [5,7].SourceTypeCfg := 1, [5,8].PVscale := 60.0, [5,8].Title := 'Phase2 CVs', [5,8].EGU := 'CVs', [5,8].EnableCfg := 1, [5,8].SourceTypeCfg := 1, [5,9].PVscale := 60.0, [5,9].Title := 'Phase3 CVs', [5,9].EGU := 'CVs', [5,9].EnableCfg := 1, [5,9].SourceTypeCfg := 1, [5,10].PVscale := 60.0, [5,10].Title := 'Phase4 CVs', [5,10].EGU := 'CVs', [5,10].EnableCfg := 1, [5,10].SourceTypeCfg := 1, [5,11].PVscale := 60.0, [5,11].Title := 'Phase5 CVs', [5,11].EGU := 'CVs', [5,11].EnableCfg := 1, [5,11].SourceTypeCfg := 1);
   PI001 : ALIAS FOR AnalogPoint[5];   // Feed Pressure
   PI001_SIG : ALIAS FOR DigitalPoint[97];
   PI001Alarm : ALIAS FOR AlarmAnalog[5];   // Feed Pressure Alarm
   PI002 : ALIAS FOR AnalogPoint[6];   // Retentate Pressure
   PI002_SIG : ALIAS FOR DigitalPoint[98];
   PI002Alarm : ALIAS FOR AlarmAnalog[6];   // Retentate Pressure Alarm
   PI101 : ALIAS FOR AnalogPoint[7];   // Filtrate Pressure
   PI101_SIG : ALIAS FOR DigitalPoint[99];
   PI101Alarm : ALIAS FOR AlarmAnalog[7];   // Filtrate Pressure Alarm
   PI401 : ALIAS FOR AnalogPoint[8];   // Transfer Pump Pressure
   PI401_SIG : ALIAS FOR DigitalPoint[100];
   PI401Alarm : ALIAS FOR AlarmAnalog[8];   // Transfer Pump Pressure Alarm
   PipeAnimation : PipeAnimation := (PipeStatP1[27] := 1, PipeStatP1[28] := 1, PipeStatP1[29] := 1, PipeStatP1[30] := 1, PipeStatP1[31] := 1, PipeStatP1[32] := 1, PipeStatP1[33] := 1, PipeStatP1[34] := 1, PipeStatP1[35] := 1, PipeStatP1[36] := 1, PipeStatP1[40] := 1, PipeStatP1[41] := 1, PipeStatP1[42] := 1, PipeStatP1[43] := 1, PipeStatP1[44] := 1, PipeStatP1[45] := 1, PipeStatP1[46] := 1, PipeStatP1[47] := 1, PipeStatP1[50] := 1, PipeStatP1[51] := 1, PipeStatP1[55] := 1, PipeStatP1[56] := 1, PipeStatP2[1] := 1, PipeStatP2[20] := 1, PipeStatP2[21] := 1, PipeStatP2[22] := 1, PipeStatP2[23] := 1, PipeStatP2[24] := 1, PipeStatP2[25] := 1, PipeStatP2[26] := 1, PipeStatP2[27] := 1, PipeStatP2[28] := 1, PipeStatP2[29] := 1, PipeStatP2[33] := 1, PipeStatP2[34] := 1, PipeStatP2[35] := 1, PipeStatP2[36] := 1, PipeStatP2[40] := 1, PipeStatP2[41] := 1, PipeStatP2[42] := 1, PipeStatP2[43] := 1, PipeStatP2[44] := 1, PipeStatP2[45] := 1, PipeStatP2[46] := 1, PipeStatP2[47] := 1, PipeStatP2[50] := 1, PipeStatP2[51] := 1, PipeStatP2[55] := 1, PipeStatP2[56] := 1);   // HMI Pipe Animation Array
   PipeStatValueHMI : INT[224] := ([1] := 1, [20] := 1, [21] := 1, [22] := 1, [23] := 1, [24] := 1, [25] := 1, [26] := 1, [27] := 1, [28] := 1, [29] := 1, [30] := 1, [31] := 1, [32] := 1, [33] := 1, [34] := 1, [35] := 1, [36] := 1, [40] := 1, [41] := 1, [42] := 1, [43] := 1, [44] := 1, [45] := 1, [46] := 1, [47] := 1, [50] := 1, [51] := 1, [55] := 1, [56] := 1);   // Pipe Animation Value For HMI
   PLCFault : FaultRecordType := (Info[0] := 3, Info[1] := 22820, Info[2] := 9248, Info[3] := 1637339701);   // PLC Major Fault Record
        .Info   // Fault specific information
        .Code   // Unique code for the fault
        .TimeLow   // Lower 32 bits of the fault timestamp value
        .TimeHigh   // Upper 32 bits of the fault timestamp value
        .RecType   // Fault Type
   ProcedureTime : ALIAS FOR Timers[19];   // Procedure Time
   Prompt : Prompt[7] := ([1].Step := 3, [1].Value := 1, [2].Step := 4, [2].Value := 1, [6].Step := 5);   // Prompt Array
   Prompt0 : ALIAS FOR Prompt[0];   // Phase 0 Prompt
   Prompt1 : ALIAS FOR Prompt[1];   // Phase 1 Prompt
   Prompt2 : ALIAS FOR Prompt[2];   // Phase 2 Prompt
   Prompt3 : ALIAS FOR Prompt[3];   // Phase 3 Prompt
   Prompt4 : ALIAS FOR Prompt[4];   // Phase 4 Prompt
   Prompt5 : ALIAS FOR Prompt[5];   // Phase 5 Prompt
   PromptTimer : FBD_TIMER := (PRE := 1000, EN := 1);   // Prompt Timer
   PSH001 : ALIAS FOR DigitalPoint[4];   // Feed Pump High Pressure
   PSH401 : ALIAS FOR DigitalPoint[5];   // Transfer Pump High Pressure
   PSL602 : ALIAS FOR DigitalPoint[0];   // Valves Air Defect
   PSL603 : ALIAS FOR DigitalPoint[10];   // Manifold Valves Air Defect
   PumpRunStatus : DINT;   // Pumps Run Status (1 = At least one pump running , 0 = no pump running)
   Rack_Murr_Node0_Smart : IO_Station := (Node_Comm_Status_value := 16384, Node_Comm_Status := 1, Node_Internal_Defect_Status := 1);   // Status of Node 0 Smart
   Rack_Murr_Node1_TF2S : IO_Station := (Node_Comm_Status_value := 24576, Node_Internal_Defect_Status := 1, Inhibition := 4);   // Status of Node 1 TF2S
   Rack_Murr_Node1_TF3S : IO_Station := (Node_Comm_Status_value := 16384, Node_Comm_Status := 1, Node_Internal_Defect_Status := 1);   // Status of Node 1 TF3S
   Rack_Murr_Node3_PUMP : IO_Station := (Node_Comm_Status_value := 16384, Node_Comm_Status := 1, Node_Internal_Defect_Status := 1);   // Status of Node 3 Pump
   Rack_Murr_Node4_Instrum_TFF1 : IO_Station := (Node_Comm_Status_value := 24576, Node_Internal_Defect_Status := 1, Inhibition := 4);   // Status of Node 4 Instrum TFF1
   Rack_Murr_Node4_Instrum_TFF2 : IO_Station := (Node_Comm_Status_value := 24576, Node_Internal_Defect_Status := 1, Inhibition := 4);   // Status of Node 4 Instrum TFF2
   Rack_Murr_Node4_Instrum_TFF3 : IO_Station := (Node_Comm_Status_value := 16384, Node_Comm_Status := 1, Node_Internal_Defect_Status := 1);   // Status of Node 4 Instrum TFF3
   Rack_Murr_Node4_Instrum_TFF4 : IO_Station := (Node_Comm_Status_value := 24576, Node_Internal_Defect_Status := 1, Inhibition := 4);   // Status of Node 4 Instrum TFF4
   Rack_Murr_Node4_Instrum_TFF5 : IO_Station := (Node_Comm_Status_value := 24576, Node_Internal_Defect_Status := 1, Inhibition := 4);   // Status of Node 4 Instrum TFF5
   Rack_Murr_Node5_Tank100 : IO_Station := (Node_Comm_Status_value := 24576, Node_Internal_Defect_Status := 1, Inhibition := 4);   // Status of Node 5 Tank 100L
   Rack_Murr_Node5_Tank250 : IO_Station := (Node_Comm_Status_value := 16384, Node_Comm_Status := 1, Node_Internal_Defect_Status_value := -53, Node_Internal_Defect_Status := 1);   // Status of Node 5 Tank 250L
   Rack_Murr_Node5_Tank50 : IO_Station := (Node_Comm_Status_value := 24576, Node_Internal_Defect_Status := 1, Inhibition := 4);   // Status of Node 5 Tank 50L
   Rack_Murr_Node6_IND331_WI001 : IO_Station := (Node_Comm_Status_value := 16384, Node_Comm_Status := 1, Node_Internal_Defect_Status := 1);   // Status of Node 6 IND331 WI001
   Rack_Murr_Node7_IND131_WI101 : IO_Station := (Node_Comm_Status_value := 16384, Node_Comm_Status := 1, Node_Internal_Defect_Status := 1);   // Status of Node 7 IND131 WI101
   RawAnalogInputArray : INT[50] := ([3] := 23481, [4] := 23321, [5] := 6540, [6] := 6482, [7] := 6484, [8] := 6656, [10] := 6559, [11] := 7802, [12] := 6960, [13] := 16334, [14] := 42, [37] := 6414);   // Array of analog input raw
   RecipeStepLog_DateTime : STRING25;
   ScaleFiltering : ScaleFiltering := (CurrentFilter := 2, Sample_Rate := 10, Timer.PRE := 99999999, Timer.EN := 1, Timer.TT := 1, FeedBagVolume_MAVE.SampleEnable := 1, FeedBagVolume_MAVE.NumberOfSamples := 1, FiltrateFlow := 0.34332275, FiltrateFlow_MAVE.In := 61.307632, FiltrateFlow_MAVE.SampleEnable := 1, FiltrateFlow_MAVE.NumberOfSamples := 1, FiltrateFlow_MAVE.Out := 61.307632, FiltrateFlow_Mave_Timer.PRE := 99999999, FiltrateFlow_Mave_Timer.EN := 1, FiltrateFlow_Mave_Timer.TT := 1, FiltrateFlow_Mave_Sample_Rate := 100, FiltrateFlow_ExpConst := 0.99, FiltrateFlow_Exp_Timer.PRE := 99999999, FiltrateFlow_Exp_Timer.ACC := 100, FiltrateFlow_Exp_Timer.EN := 1, FiltrateFlow_Exp_Timer.TT := 1, FiltrateFlow_Exp_Sample_Rate := 100, FiltrateFlow_ExpFiltered := -0.0011392268, FiltrateVolume101_MAVE.SampleEnable := 1, FiltrateVolume101_MAVE.NumberOfSamples := 1, FiltrateVolume101_ExpConst := 0.99, WI102_Unfiltered := -374.97137, FiltrateVolume102 := -374.97137, FiltrateVolume102_Array[0] := -374.91415, FiltrateVolume102_Array[1] := -374.97137, FiltrateVolume102_Array[2] := -374.97137, FiltrateVolume102_Array[3] := -374.97137, FiltrateVolume102_Array[4] := -374.97137, FiltrateVolume102_Array[5] := -374.91415, FiltrateVolume102_Array[6] := -374.91415, FiltrateVolume102_Array[7] := -374.97137, FiltrateVolume102_Array[8] := -374.97137, FiltrateVolume102_Array[9] := -374.97137, FiltrateVolume102_Array[10] := -374.97137, FiltrateVolume102_Array[11] := -374.97137, FiltrateVolume102_Array[12] := -374.97137, FiltrateVolume102_Array[13] := -374.97137, FiltrateVolume102_Array[14] := -374.97137, FiltrateVolume102_Array[15] := -374.97137, FiltrateVolume102_Array[16] := -374.97137, FiltrateVolume102_Array[17] := -374.97137, FiltrateVolume102_Array[18] := -374.97137, FiltrateVolume102_Array[19] := -374.97137, FiltrateVolume102_Array[20] := -374.97137, FiltrateVolume102_Array[21] := -374.97137, FiltrateVolume102_Array[22] := -374.97137, FiltrateVolume102_Array[23] := -374.97137, FiltrateVolume102_Array[24] := -374.97137, FiltrateVolume102_Array[25] := -374.97137, FiltrateVolume102_Array[26] := -374.91415, FiltrateVolume102_Array[27] := -374.97137, FiltrateVolume102_Array[28] := -374.97137, FiltrateVolume102_Array[29] := -374.91415, FiltrateVolume102_Array[30] := -374.97137, FiltrateVolume102_Array[31] := -374.97137,
        FiltrateVolume102_Array[32] := -374.97137, FiltrateVolume102_Array[33] := -374.85693, FiltrateVolume102_Array[34] := -374.97137, FiltrateVolume102_Array[35] := -374.97137, FiltrateVolume102_Array[36] := -374.97137, FiltrateVolume102_Array[37] := -374.97137, FiltrateVolume102_Array[38] := -374.91415, FiltrateVolume102_Array[39] := -374.97137, FiltrateVolume102_Array[40] := -374.85693, FiltrateVolume102_Array[41] := -374.97137, FiltrateVolume102_Array[42] := -374.97137, FiltrateVolume102_Array[43] := -374.97137, FiltrateVolume102_Array[44] := -374.97137, FiltrateVolume102_Array[45] := -374.97137, FiltrateVolume102_Array[46] := -374.91415, FiltrateVolume102_Array[47] := -374.97137, FiltrateVolume102_Array[48] := -374.97137, FiltrateVolume102_Array[49] := -374.91415, FiltrateVolume102_Array[50] := -374.97137, FiltrateVolume102_Array[51] := -374.97137, FiltrateVolume102_Array[52] := -374.85693, FiltrateVolume102_Array[53] := -374.97137, FiltrateVolume102_Array[54] := -374.85693, FiltrateVolume102_Array[55] := -374.97137, FiltrateVolume102_Array[56] := -374.97137, FiltrateVolume102_Array[57] := -374.91415, FiltrateVolume102_Array[58] := -374.97137, FiltrateVolume102_Array[59] := -374.97137, FiltrateVolume102_Array[60] := -374.97137, FiltrateVolume102_Array[61] := -374.97137, FiltrateVolume102_Array[62] := -374.97137, FiltrateVolume102_Array[63] := -374.97137, FiltrateVolume102_Array[64] := -374.97137, FiltrateVolume102_Array[65] := -374.97137, FiltrateVolume102_Array[66] := -374.97137, FiltrateVolume102_Array[67] := -374.97137, FiltrateVolume102_Array[68] := -374.97137, FiltrateVolume102_Array[69] := -374.97137, FiltrateVolume102_Array[70] := -374.97137, FiltrateVolume102_Array[71] := -374.97137, FiltrateVolume102_Array[72] := -374.97137, FiltrateVolume102_Array[73] := -374.97137, FiltrateVolume102_Array[74] := -374.97137, FiltrateVolume102_Array[75] := -374.97137, FiltrateVolume102_Array[76] := -374.97137, FiltrateVolume102_Array[77] := -374.97137, FiltrateVolume102_Array[78] := -374.97137, FiltrateVolume102_Array[79] := -374.97137, FiltrateVolume102_Array[80] := -374.97137, FiltrateVolume102_Array[81] := -374.97137, FiltrateVolume102_Array[82] := -374.97137, FiltrateVolume102_Array[83] := -374.91415, FiltrateVolume102_Array[84] := -374.97137, FiltrateVolume102_Array[85] := -374.97137, FiltrateVolume102_Array[86] := -374.97137, FiltrateVolume102_Array[87] := -374.91415, FiltrateVolume102_Array[88] := -374.97137, FiltrateVolume102_Array[89] := -374.97137, FiltrateVolume102_Array[90] := -374.97137, FiltrateVolume102_Array[91] := -374.91415,
        FiltrateVolume102_Array[92] := -374.97137, FiltrateVolume102_Array[93] := -374.97137, FiltrateVolume102_Array[94] := -374.97137, FiltrateVolume102_Array[95] := -374.97137, FiltrateVolume102_Array[96] := -374.97137, FiltrateVolume102_Array[97] := -374.97137, FiltrateVolume102_Array[98] := -374.91415, FiltrateVolume102_Array[99] := -374.91415, FiltrateVolume102_Array[100] := -374.97137, FiltrateVolume102_MAVE.In := -374.97137, FiltrateVolume102_MAVE.SampleEnable := 1, FiltrateVolume102_MAVE.NumberOfSamples := 1, FiltrateVolume102_MAVE.Out := -374.97137, FiltrateVolume102_MaveFiltered := -374.97137, FiltrateVolume102_ExpConst := 0.99, FiltrateVolume102_ExpFiltered := -374.9605, Weight102_ExpFiltered := -374.9605, Weight102_MaveFiltered := -374.97137, FiltrateVolume_ExpFiltered := -374.9605, FiltrateVolume_ExpFiltered_Prev := -374.96072, FiltrateVolume_MaveFiltered := -374.97137, FiltrateVolume_MaveFiltered_Prev := -374.85693);   // Data for Scale Filtering
   SIC001 : ALIAS FOR Drive[1];   // Feed Pump
   SIC001_AO : ALIAS FOR AnalogOutput[2];   // Feed Pump Speed Setpoint
   SIC001DF : ALIAS FOR DigitalPoint[8];   // Feed Pump Defect
   SIC002 : ALIAS FOR Drive[2];   // Transfer Pump
   SIC002_AO : ALIAS FOR AnalogOutput[3];   // Transfer Pump Speed Setpoint
   SIC002DF : ALIAS FOR DigitalPoint[9];   // Transfer Pump Defect
   SIC003 : ALIAS FOR Drive[3];   // Mixer
   SIC003_AO : ALIAS FOR AnalogOutput[4];   // Mixer Speed Setpoint
   SIC003DF : ALIAS FOR DigitalPoint[14];   // Mixer Defect
   SRL001 : ALIAS FOR DigitalPoint[15];   // Tank Skid Remote / Standalone
   SysControl : SysControl := (DefaultTimer.PRE := 3000, AllAutoTimer.PRE := 3000, DefaultStatus := 1, UV_Auto_Zero_Timer.PRE := 3000);   // General system status and command
   Tank : TankManagement := (Config.TankSelected := 3, Config.TankSelectHMI := 3, Config.Option_Current := 3, Config.Option_Prev := 3, Config.TMR.PRE := 500, Config.AlarmStatus := 1, WeightConfiguration[0].Alm_HI := 2.0, WeightConfiguration[0].Alm_HI_PRE := 2.0, WeightConfiguration[0].Alm_HIHI := 2.0, WeightConfiguration[0].Alm_HIHI_PRE := 2.0, WeightConfiguration[0].Alm_LOLOTMR := 2, WeightConfiguration[0].Alm_LOLOTMR_PRE := 2, WeightConfiguration[0].Alm_LOTMR := 2, WeightConfiguration[0].Alm_LOTMR_PRE := 2, WeightConfiguration[0].Alm_HITMR := 2, WeightConfiguration[0].Alm_HITMR_PRE := 2, WeightConfiguration[0].Alm_HIHITMR := 2, WeightConfiguration[0].Alm_HIHITMR_PRE := 2, WeightConfiguration[1].Alm_HI := 60.0, WeightConfiguration[1].Alm_HI_PRE := 60.0, WeightConfiguration[1].Alm_HIHI := 60.0, WeightConfiguration[1].Alm_HIHI_PRE := 60.0, WeightConfiguration[1].Alm_LOLOTMR := 2, WeightConfiguration[1].Alm_LOLOTMR_PRE := 2, WeightConfiguration[1].Alm_LOTMR := 2, WeightConfiguration[1].Alm_LOTMR_PRE := 2, WeightConfiguration[1].Alm_HITMR := 2, WeightConfiguration[1].Alm_HITMR_PRE := 2, WeightConfiguration[1].Alm_HIHITMR := 2, WeightConfiguration[1].Alm_HIHITMR_PRE := 2, WeightConfiguration[2].Alm_LOLO := 99.999, WeightConfiguration[2].Alm_LOLO_PRE := 99.999, WeightConfiguration[2].Alm_LO := 199.998, WeightConfiguration[2].Alm_LO_PRE := 199.998, WeightConfiguration[2].Alm_HI := 799.992, WeightConfiguration[2].Alm_HI_PRE := 799.992, WeightConfiguration[2].Alm_HIHI := 899.99097, WeightConfiguration[2].Alm_HIHI_PRE := 899.99097, WeightConfiguration[2].Alm_LOLOTMR := 2, WeightConfiguration[2].Alm_LOLOTMR_PRE := 2, WeightConfiguration[2].Alm_LOTMR := 2, WeightConfiguration[2].Alm_LOTMR_PRE := 2, WeightConfiguration[2].Alm_HITMR := 2, WeightConfiguration[2].Alm_HITMR_PRE := 2, WeightConfiguration[2].Alm_HIHITMR := 2, WeightConfiguration[2].Alm_HIHITMR_PRE := 2, WeightConfiguration[3].Alm_HI := 230.0, WeightConfiguration[3].Alm_HI_PRE := 230.0, WeightConfiguration[3].Alm_HIHI := 240.0, WeightConfiguration[3].Alm_HIHI_PRE := 240.0, LevelConfiguration[0].Alm_HI := 99999.0, LevelConfiguration[0].Alm_HI_PRE := 99999.0, LevelConfiguration[0].Alm_HIHI := 99999.0, LevelConfiguration[0].Alm_HIHI_PRE := 99999.0, LevelConfiguration[0].Alm_LOLOTMR := 2, LevelConfiguration[0].Alm_LOLOTMR_PRE := 2, LevelConfiguration[0].Alm_LOTMR := 2, LevelConfiguration[0].Alm_LOTMR_PRE := 2, LevelConfiguration[0].Alm_HITMR := 2, LevelConfiguration[0].Alm_HITMR_PRE := 2,
